(* IEC 61131-3 sources: daoli-st-library/DL_MathData (part 22) *)

(* ---- FC_DL_RealToUintSat.st ---- *)
(*
    FC_DL_RealToUintSat —— REAL 到 UINT 饱和防御转换
    ------------------------------------------------------------------
    分类      : DL_MathData / Convert
    前缀      : FC_DL_
    版本      : 1.0.0
    溯源      : IEC 61131-3 标准语义的道莅防御性实现
                （内部委托平台内建函数，外围统一错误码/钳位/双语文档；
                  未复制任何闭源厂商源码，参考实现仅限 MIT/Apache 许可）
    平台      : 纯 IEC 61131-3，CODESYS / TwinCAT / InoProShop 通用
    作者      : 道莅代码库 · PLC编程专家（R16）
    ------------------------------------------------------------------
    功能说明  : 将 REAL 输入防御性转换为 UINT 并作为返回值输出；
                非有限输入（NaN 或 ±INF）判为故障级 16#0001_0297，返回 0 且 bValid=FALSE；
                fIn < 0 时钳位至 0，置信息级 16#0001_01C6（UINT 无符号，负值不可表）；
                fIn 超出 UINT 上界 65535 时钳位至上界，置信息级 16#0001_01C7；
                钳位方向：下界 0 / 上界 65535（双侧饱和）；
                ±INF 采用平台安全幅值比较判定（阈值高于 REAL 最大有限值 3.402823E38），NaN 用 fIn <> fIn 自不等判定；
                域内转换委托平台内建 REAL_TO_UINT 语义，不重实现数学内核；
                信息级码属正常防御：bError=FALSE、bValid=TRUE，输出钳位后防御值。
    错误码    : 16#0001_0297 非有限输入（NaN 或 ±INF）——故障级，返回 0
                16#0001_01C6 负值输入，已钳位至 0——信息级，正常防御
                16#0001_01C7 输入超 UINT 上界，已钳位至 65535——信息级，正常防御
                16#0001_0298 预留禁用（故障级，不得挪用）
                16#0001_0299 预留禁用（故障级，不得挪用）
    状态机    : R6 标注 N/A —— 本组件为纯函数无顺序状态机，无 CASE 可写，非法状态不可能出现，故以本节说明替代 ELSE 兜底
    修订记录  : 2026-11-16 v1.0.0 首次入库（R16）
*)
FUNCTION FC_DL_RealToUintSat : UINT
VAR_INPUT
    fIn : REAL; // 待转换输入 [无量纲] / input value to convert
END_VAR
VAR_OUTPUT
    eErr   : UDINT; // 错误码，0=正常 / error id, 0=ok
    bError : BOOL;  // 是否出错，eErr 非 0 时为 TRUE / error flag, TRUE when eErr is nonzero
    bValid : BOOL;  // 输出是否有效可用 / output valid flag
END_VAR
VAR CONSTANT
    DL_UINT16_MAX     : LREAL := 65535.0; // UINT 域上界 65535，LREAL 承载 [无量纲] / UINT upper bound 65535 carried in LREAL
    DL_REAL_INF_GUARD : LREAL := 4.0E38;  // REAL 域 ±INF 判定阈值，高于 REAL 最大有限值 3.402823E38 [无量纲] / REAL +/-INF guard above max finite REAL 3.402823E38
END_VAR
VAR
    bNonFinite : BOOL; // 非有限（NaN 或 ±INF）判定结果 / non-finite (NaN or +/-INF) detection result
END_VAR

// 段 1｜返回值与错误状态预置 / segment 1, preset return value and error status
FC_DL_RealToUintSat := 0; // 故障缺省返回 0 [无量纲] / fault default returns 0
eErr   := 0;     // 预置无错误 / preset no error
bError := FALSE; // 预置无故障 / preset no fault
bValid := FALSE; // 预置无效，通过防御闸后置位 / preset invalid, set TRUE after guard passes

// 段 2｜非有限防御闸 / segment 2, non-finite guard
bNonFinite := (fIn <> fIn) OR (fIn > DL_REAL_INF_GUARD) OR (fIn < -DL_REAL_INF_GUARD); // NaN 自不等判定，±INF 用安全幅值比较 [无量纲] / NaN by self-inequality, +/-INF by safe magnitude compare
IF bNonFinite THEN
    FC_DL_RealToUintSat := 0; // 故障级返回 0 [无量纲] / fault level returns 0
    eErr   := 16#0001_0297;   // 非有限输入故障码 / non-finite input fault id
    bError := TRUE;           // 置故障标志 / set fault flag
    bValid := FALSE;          // 输出无效 / output invalid
    RETURN;                   // 立即返回 / immediate return
END_IF

// 段 3｜双侧饱和钳位与主体转换（末段） / segment 3, double-side saturating clamp and main conversion (final)
IF fIn < 0.0 THEN
    FC_DL_RealToUintSat := 0;  // 负值钳位至 0（UINT 无符号语义） / negative input clamped to 0 (UINT is unsigned)
    eErr := 16#0001_01C6;      // 信息级：负值已钳零 / info level: negative input clamped to zero
ELSIF fIn > DL_UINT16_MAX THEN
    FC_DL_RealToUintSat := 16#FFFF; // 正向钳位至 UINT 上界 65535 / clamp to UINT upper bound 65535
    eErr := 16#0001_01C7;           // 信息级：超上界已钳位 / info level: above upper bound, clamped
ELSE
    FC_DL_RealToUintSat := REAL_TO_UINT(fIn); // 域内委托平台内建 _TO_ 转换语义 / in-domain delegate to built-in _TO_ conversion
    eErr := 0; // 域内无错误 / in-domain, no error
END_IF
bError := FALSE; // 信息级钳位不置故障，故障分支已提前返回 / info-level clamp never raises fault, fault branch has returned
bValid := TRUE;  // 域内或钳位输出均有效可用 / in-domain or clamped output is valid
END_FUNCTION

(* ---- FC_DL_ReverseBitsWord.st ---- *)
(*==============================================================================
 * 组件名称 (Component)  : FC_DL_ReverseBitsWord
 * 所属子库 (Sublibrary) : DL_MathData
 * 归属目录 (Directory)  : C:\Library\DL_MathData
 * 当前版本 (Version)    : 1.0.0
 * 分类/来源标签         : 函数（FUNCTION）· 纯函数 · WORD 位反转与字节交换
 *                         iec-std-wrapper / bitstring
 * 兼容性   (Platform)   : CODESYS 3.5 / TwinCAT 3 / 汇川 InoProShop / 施耐德
 *                         Machine Expert；仅用 IEC 标准位运算 AND/OR/SHL/SHR
 * 溯源声明 (Provenance) : IEC 61131-3 标准语义的道莅防御性实现——内部委托平台标准库语义，
 *                         外围统一错误码 / 钳位 / 双语注释，严禁重实现数学内核。
 * 功能一句话 (Summary)  : WORD 全 16 位镜像反转（分治交换法）或字节序交换双模式，
 *                         服务 LSB-first CRC、LED 点阵与大小端报文适配。
 *
 * 功能描述 (Function)   : 位反转模式用四步分治交换（1 位组、2 位组、4 位组、
 *                         8 位组两两对换）实现全位镜像，无循环、无查表、常数时间；
 *                         字节交换模式一次完成高低字节对换；模式域外走 ELSE 兜底
 *                         回退位反转并报故障码，回文输入以信息级告知恒等结果。
 * 与既有件边界 (Boundary): 与 ShlEx/ShrEx 族正交——那些件做移位，本件做镜像；
 *                         平台内建 SWAP 指令非 IEC 标准，故字节交换同样手写实现。
 * 码位说明 (Codes)      : 信息 16#0002_3044 反转完成且结果回文（wOut 等于 wIn）
 *                         故障 16#0002_3045 模式域外，已回退位反转并照常输出
 *                         段 16#02_3_44~47，本件实占 44~45 两码。
 * 依赖说明 (Depends)    : 无 DL_ 内部依赖；零库函数依赖，纯 IEC 位运算符。
 * 红线自检 (Redline)    : 零全局依赖 ｜ 零 VAR_EXTERNAL ｜ 零 %I/%Q ｜ 纯 IEC 位运算
 *                         移位量 1/2/4/8 恒小于 16 位宽（归一达标）｜ 无除法面
 *                         ENUM 配 CASE 且 ELSE 兜底 ｜ 全变量双语同行注释
 * 修订历史 (Revision)   : 2026-11-18  v1.0.0  首版入库（R32 · 批 1）
 *============================================================================*)

FUNCTION FC_DL_ReverseBitsWord : BOOL
VAR_INPUT
    wIn   : WORD;                       // 源字 [位串] / Source word
    eMode : (eRevBits := 0, eRevBytes := 1);    // 模式枚举：全位反转或字节交换 / Mode enum: full bit reverse or byte swap
END_VAR
VAR_OUTPUT
    wOut    : WORD;                     // 反转结果 [位串] / Reversed result
    bPalin  : BOOL;                     // 回文标志，wOut 等于 wIn 时为真 / TRUE when the result equals the input
    uErrorId: UDINT;                    // 事件码，0 表示无事件 / Event code, zero means none
END_VAR
VAR
    w1 : WORD;    // 第一步交换结果（1 位组）[位串] / Stage one result, one-bit groups
    w2 : WORD;    // 第二步交换结果（2 位组）[位串] / Stage two result, two-bit groups
    w3 : WORD;    // 第三步交换结果（4 位组）[位串] / Stage three result, four-bit groups
    w4 : WORD;    // 第四步交换结果（8 位组，即全镜像）[位串] / Stage four result, full mirror
    uCode : UDINT; // 码位暂存，出口单点写入 [码] / Code staging
END_VAR

(* 段 1｜输出预置 / Pre-set *)
FC_DL_ReverseBitsWord := FALSE;
wOut    := 16#0000;
bPalin  := FALSE;
uErrorId := 16#0000_0000;
uCode   := 16#0000_0000;

(* 段 2｜模式分派（ENUM 配 CASE，ELSE 兜底拦截域外值）/ Mode dispatch with ELSE interception *)
CASE eMode OF

    eRevBits:
        (* 四步分治交换：相邻 1 位、2 位、4 位对换，最后高低 8 位整体对换
         * Four divide-and-conquer stages, constant time, no loop and no table *)
        w1 := ((wIn  AND 16#5555) SHL 1)  OR ((wIn  AND 16#AAAA) SHR 1);  // 相邻 1 位对换 / Adjacent one-bit swap
        w2 := ((w1   AND 16#3333) SHL 2)  OR ((w1   AND 16#CCCC) SHR 2);  // 相邻 2 位对换 / Adjacent two-bit swap
        w3 := ((w2   AND 16#0F0F) SHL 4)  OR ((w2   AND 16#F0F0) SHR 4);  // 相邻 4 位对换 / Adjacent four-bit swap
        w4 := ((w3   AND 16#00FF) SHL 8)  OR ((w3   AND 16#FF00) SHR 8);  // 高低 8 位对换，完成全镜像 / Final mirror
        wOut := w4;

    eRevBytes:
        (* 字节交换：低 8 位左移到高位，高 8 位右移到低位 / Swap the two bytes *)
        wOut := ((wIn AND 16#00FF) SHL 8) OR ((wIn AND 16#FF00) SHR 8);

ELSE
    (* 域外兜底：枚举被非法赋值（如强转越界）时回退位反转，绝不输出未定义值
     * Out-of-domain fallback: revert to bit reverse, never output an undefined value *)
    w1 := ((wIn  AND 16#5555) SHL 1)  OR ((wIn  AND 16#AAAA) SHR 1);
    w2 := ((w1   AND 16#3333) SHL 2)  OR ((w1   AND 16#CCCC) SHR 2);
    w3 := ((w2   AND 16#0F0F) SHL 4)  OR ((w2   AND 16#F0F0) SHR 4);
    w4 := ((w3   AND 16#00FF) SHL 8)  OR ((w3   AND 16#FF00) SHR 8);
    wOut := w4;
    uCode := 16#0002_3045;           // 故障级：模式域外已回退 / Fault: mode out of domain, reverted

END_CASE

(* 段 3｜回文告知与出口 / Palindrome notice and exit *)
IF wOut = wIn THEN
    bPalin := TRUE;                  // 恒等结果（回文字）告知 / Inform the identity result
    IF uCode = 16#0000_0000 THEN
        uCode := 16#0002_3044;       // 信息级：结果回文 / Info: palindromic result
    END_IF
END_IF
uErrorId := uCode;                   // 码位单点写入 / Single write point for the code
FC_DL_ReverseBitsWord := TRUE;
END_FUNCTION

(* ---- FC_DL_RmsCalc.st ---- *)
(*
    FC_DL_RmsCalc —— 窗口均方根（增量式平方累加防溢出 + 窗长钳位 + 非有限剔除）
    ------------------------------------------------------------------
    分类      : DL_MathData / Math-Statistics
    前缀      : FC_DL_
    版本      : 1.0.1
    来源标签  : iec-std-wrapper（T0）
    溯源      : IEC 61131-3 标准语义的道莅防御性实现
                （无状态纯函数，SQRT 为 IEC 标准内建；未复制任何闭源厂商源码）
    平台      : 纯 IEC 61131-3，CODESYS / TwinCAT / InoProShop 通用
    分工声明  : 与存量 FB_DL_SignalStatistics / FC_DL_StdDevOnline 分工——
                SignalStatistics 为驻留统计族（均值/方差多出口），StdDevOnline
                为在线流式标准差；本件为无状态数组窗口 RMS 单出口口径，
                与批 2 Safe 族惯性一致（无依赖，仅排期顺延）。
    作者      : 道莅代码库 · PLC 编程专家（R57）
    ------------------------------------------------------------------
    功能说明  : 对输入数组前 nCount 个样本求均方根。增量式累加 sum += x²/n
                防大数平方溢出（先除后加，边界十二）；窗长钳位 1..4096；
                非有限样本剔除并计数出口；有效样本数为零判错误返回 0。
    错误码    : 0000 正常 / 16#0003_0003 窗长已钳位 / 16#0003_0004 有效样本为零
                / 16#0003_0005 非有限样本已剔除（信息级，bValid 保持 TRUE）
    bValid 偏离段: 部分剔除时 bValid 保持 TRUE——有效样本统计量仍可用（与
                0303 钳位件 bValid=FALSE 的口径差异在此声明，v1.0.1）。
    修订记录  : 2026-11-21 v1.0.0 首次入库（R57 批 3 · 序号 12）
                2026-11-21 v1.0.1 R58 返修：部分剔除（nUsed>0 且 nNanCnt>0）
                置信息级 0003_0005（首事件闸），调用方可感知口径已收窄；
                全剔除路径 0304 优先级在先不动。
*)
FUNCTION FC_DL_RmsCalc : LREAL
VAR_IN_OUT
    afData : ARRAY[0..4095] OF LREAL; // 样本数组 [工程单位]，前 nCount 个有效 / the sample array, the first nCount entries valid
END_VAR
VAR_INPUT
    nCount : DINT; // 样本数 [个]，钳位 1..4096 / the sample count, clamped to one through four thousand ninety six
END_VAR
VAR_OUTPUT
    eErr     : UDINT; // 错误码，0 = 正常 / error code, zero is ok
    bError   : BOOL;  // 出错标志，eErr 非 0 时为真 / error flag, true when eErr is nonzero
    bValid   : BOOL;  // 结果是否为真实值，钳位/剔除降级时可能为假 / the result is the true value, false when degraded
    nNanCnt  : UDINT; // 剔除的非有限样本数 [个] / the excluded non finite sample count
END_VAR
VAR
    nI     : DINT;  // 循环计数 [个] / the loop counter
    nUsed  : DINT;  // 实际参与样本数 [个] / the actually used sample count
    lrSum  : LREAL; // 增量式平方和 [工程单位平方] / the incremental sum of squares
    lrX    : LREAL; // 当前样本 [工程单位] / the current sample [engineering unit]
    bClamp : BOOL;  // 窗长钳位发生 [-] / a window clamp happened
END_VAR
VAR CONSTANT
    DL_RMS_NMAX : DINT := 4096; // 窗长上限 [个]，与数组容量一致 / the window bound, aligned with the array capacity
END_VAR

// 段 1｜返回值与错误状态预置安全值（四段式第一段，R45）/ segment 1, preset the return and error states
FC_DL_RmsCalc := 0.0; // 返回值预置安全值 0.0 / preset the return to the safe zero
eErr   := 16#0000_0000; // 错误码预置正常 / preset the code to ok
bError := FALSE; // 错误标志预置假 / preset the error flag false
bValid := TRUE; // 有效标志预置真 / preset the valid flag true
nNanCnt := 0; // 剔除计数预置零 / preset the excluded count zero
bClamp := FALSE; // 钳位标志预置假 / preset the clamp flag false

// 段 2｜窗长钳位 1..4096（边界十二；上界与数组容量一致，索引结构性安全）/ segment 2, the window clamp
IF nCount < 1 THEN // 低于下界 / below the floor
    nCount := 1; // 钳到 1 / clamp to one
    bClamp := TRUE; // 置钳位标记 / raise the clamp flag
ELSIF nCount > DL_RMS_NMAX THEN // 高于上界 / above the bound
    nCount := DL_RMS_NMAX; // 钳到上限 / clamp to the bound
    bClamp := TRUE; // 置钳位标记 / raise the clamp flag
END_IF
IF bClamp THEN // 钳位发生时置信息级 / raise the informational code on a clamp
    eErr   := 16#0003_0003; // 信息级：窗长已钳位 / informational, the window clamped
    bError := TRUE; // 置错误标志 / raise the error flag
    bValid := FALSE; // 钳位口径非原始窗长口径 / the clamped window is not the requested one
END_IF

// 段 3｜增量式平方累加：sum += x²/n（先除后加防大数溢出，边界十二）/ segment 3, the incremental accumulation
lrSum := 0.0; // 平方和清零 / clear the sum
nUsed := 0; // 参与样本数清零 / clear the used count
FOR nI := 0 TO nCount - 1 DO // 有界循环（nCount 已钳 ≤4096）/ the bounded loop
    lrX := afData[nI]; // 取样本（索引已证在数组界内）/ take the sample, the index proven inside the bounds
    IF (lrX = lrX) AND ((lrX - lrX) = (lrX - lrX)) THEN // 非有限双判据通过才参与 / only finite samples participate
        lrSum := lrSum + lrX * lrX / INT_TO_LREAL(nCount); // 先除窗长再加，防 x² 大数溢出 / divide first then add against overflow
        nUsed := nUsed + 1; // 参与计数推进 / advance the used count
    ELSE // 非有限样本剔除 / a non finite sample excluded
        nNanCnt := nNanCnt + 1; // 剔除计数推进 / advance the excluded count
    END_IF
END_FOR

// 段 3b｜部分剔除信息级置码（v1.0.1：首事件闸，0303 先发则不再覆盖）/ segment 3b, the partial exclusion informational code
IF (nNanCnt > 0) AND (nUsed > 0) AND (eErr = 16#0000_0000) THEN // 部分剔除且无先发事件 / a partial exclusion with no earlier event
    eErr   := 16#0003_0005; // 信息级：非有限样本已剔除，口径为有效样本 RMS / informational, non finite samples excluded, the effective sample RMS
    bError := TRUE; // 置错误标志（信息级随事件置位惯例）/ raise the error flag
END_IF // bValid 保持 TRUE：有效样本统计量仍可用（头注释偏离段声明）/ bValid stays true, the effective sample statistic remains usable

// 段 4｜结果计算与兜底 / segment 4, the result and the guard
IF nUsed > 0 THEN // 有有效样本 / with valid samples
    FC_DL_RmsCalc := SQRT(lrSum * INT_TO_LREAL(nCount) / INT_TO_LREAL(nUsed)); // 复原除子后开方（除子已证大于零）/ restore the divisor then the square root
ELSE // 全部剔除 / all excluded
    eErr   := 16#0003_0004; // 错误级：有效样本为零 / error grade, no valid sample
    bError := TRUE; // 置错误标志 / raise the error flag
    bValid := FALSE; // 输出不可用 / the output void
END_IF
IF (FC_DL_RmsCalc <> FC_DL_RmsCalc) OR ((FC_DL_RmsCalc - FC_DL_RmsCalc) <> (FC_DL_RmsCalc - FC_DL_RmsCalc)) THEN // 结果非有限兜底 / the non finite result guard
    FC_DL_RmsCalc := 0.0; // 兜底安全值 / the bottom-line safe value
    bValid := FALSE; // 输出不可用 / the output void
END_IF
END_FUNCTION

(* ---- FC_DL_RoundBankEx.st ---- *)
(*
    FC_DL_RoundBankEx —— ROUND 明确口径包装（银行家/半进可选，LREAL 域）
    ------------------------------------------------------------------
    分类      : DL_MathData / Rounding
    前缀      : FC_DL_
    版本      : 1.0.0
    溯源      : IEC 61131-3 标准语义的道莅防御性实现
                （内部委托 TRUNC 标准函数与比较语义，外围统一错误码/钳位/双语文档；
                  未复制任何闭源厂商源码，参考实现仅限 MIT/Apache 许可）
    平台      : 纯 IEC 61131-3，CODESYS / TwinCAT / InoProShop 通用
    作者      : 道莅代码库 · PLC编程专家（R40）
    ------------------------------------------------------------------
    功能说明  : 将 fIn 舍入到最近整数（仍以 LREAL 返回），0.5 进位方向全平台
                显式统一，杜绝 ROUND 内建在三平台的半进/半退差异泄漏：
                bHalfUp = FALSE（缺省）：0.5 进位到最近的偶数（银行家口径）；
                bHalfUp = TRUE：0.5 一律进位（向远离零方向，半进口径）；
                非半点小数一律按最近整数舍入（>0.5 进、<0.5 退）；
                非有限输入（NaN 或 ±Inf）判为故障级 16#0001_03CF，返回 0.0 且
                bValid=FALSE（NaN 参与舍入在三平台行为不一致，一律拦截）；
                超整数分辨率恒等直通：|fIn| ≥ 2^53（9.007199254740992E15）时
                该幅值下 LREAL 相邻可表数间距已大于 1，输入必为整数值，
                舍入恒等直通并置信息级 16#0001_0496；
                溢出面分析（R63 反算句）：|fIn| < 2^53 时结果 |fRnd| ≤ |fIn| + 1 ≤ 2^53，
                恒在 LREAL 可表域内，无溢出路径，无需饱和钳位（算法已证）；
                半点检测口径：ABS(fFrac − 0.5) < 1.0E-9 视为半点（差值在 1E-9 内的
                近半点值按半点口径处理，取舍显式化，避免浮点表示误差致半点漏判）。
    错误码    : 16#0001_03CF 任一输入非有限（NaN 或 ±Inf）——故障级，返回 0.0
                16#0001_0496 输入幅值 ≥ 2^53，超整数分辨率，恒等直通——信息级，正常防御
                （R90 反证句：恒等直通场景无法由返回值观测——直通值与舍入结果同为
                  合法整数值，bValid=TRUE 组合相同，现有输出无法还原「分辨率已耗尽」
                  事实，故占信息码）
    状态机    : R6 标注 N/A —— 本组件为纯函数无顺序状态机，无 CASE 可写，
                非法状态不可能出现，故以本节说明替代 ELSE 兜底
    修订记录  : 2026-11-19 v1.0.0 首次入库（R40 · 批 2 · T0 快车道）
*)
FUNCTION FC_DL_RoundBankEx : LREAL
VAR_INPUT
    fIn     : LREAL;         // 待舍入输入 [无量纲] ｜ input to round
    bHalfUp : BOOL := FALSE; // 半点口径，FALSE=进位到最近偶数（银行家），TRUE=一律半进 ｜ half-point mode, FALSE=round half to even (banker's), TRUE=round half away from zero
END_VAR
VAR_OUTPUT
    eErr   : UDINT; // 错误码，0=正常，16#0001_04XX=信息级，16#0001_03XX=故障级 ｜ error id, 0=ok, 16#0001_04XX=info, 16#0001_03XX=fault
    bError : BOOL;  // 是否出错，eErr 落故障级时为 TRUE ｜ fault flag, TRUE when eErr is fault level
    bValid : BOOL;  // 输出是否有效可用 ｜ output valid flag
END_VAR
VAR CONSTANT
    DL_ROUND_ID_LIMIT : LREAL := 9.007199254740992E15; // 恒等直通幅值限 = 2^53 [无量纲] ｜ identity pass-through magnitude limit = 2^53
    DL_ROUND_HALF     : LREAL := 0.5;                  // 半点判据常数 [无量纲] ｜ half-point constant
    DL_ROUND_TOL      : LREAL := 1.0E-9;               // 半点检测容差 [无量纲] ｜ half-point detection tolerance
    DL_ROUND_ONE      : LREAL := 1.0;                  // 进位步长 [无量纲] ｜ carry step
    DL_ROUND_TWO      : LREAL := 2.0;                  // 偶数判定基数 [无量纲] ｜ even-test radix
END_VAR
VAR
    bNonFinite : BOOL;  // 非有限（NaN 或 ±Inf）判定结果 ｜ non-finite (NaN or +/-Inf) detection result
    fAbs       : LREAL; // 输入绝对值 [无量纲] ｜ absolute value of the input
    fInt       : LREAL; // 绝对值的整数部分（TRUNC 向零截断）[无量纲] ｜ integer part of the magnitude (TRUNC toward zero)
    fFrac      : LREAL; // 绝对值的小数部分 [无量纲] ｜ fractional part of the magnitude
    fRnd       : LREAL; // 舍入后的绝对值结果 [无量纲] ｜ rounded magnitude result
END_VAR

// 段 1｜返回值与错误状态预置 ｜ segment 1, preset return value and error status
FC_DL_RoundBankEx := 0.0; // 故障缺省返回 0 [无量纲] ｜ fault default returns 0
eErr   := 0;     // 预置无错误 ｜ preset no error
bError := FALSE; // 预置无故障 ｜ preset no fault
bValid := FALSE; // 预置无效，通过防御闸后置位 ｜ preset invalid, set TRUE after guard passes

// 段 2｜非有限防御闸（早退） ｜ segment 2, non-finite guard (early return)
bNonFinite := (fIn <> fIn) OR ((fIn - fIn) <> (fIn - fIn)); // NaN 自不等 + 差值自减判 ±Inf [无量纲] ｜ NaN by self-inequality, +/-Inf by self-subtraction
IF bNonFinite THEN
    FC_DL_RoundBankEx := 0.0; // 故障级返回 0 [无量纲] ｜ fault level returns 0
    eErr   := 16#0001_03CF;   // 非有限输入故障码 ｜ non-finite input fault id
    bError := TRUE;           // 置故障标志（R45 配对）｜ raise the fault flag (R45 pairing)
    bValid := FALSE;          // 输出无效 ｜ output invalid
    RETURN;                   // 早退 ｜ early return
END_IF

// 段 3｜超整数分辨率恒等直通（信息级） ｜ segment 3, identity pass-through beyond integer resolution (info level)
IF ABS(fIn) >= DL_ROUND_ID_LIMIT THEN
    FC_DL_RoundBankEx := fIn; // 分辨率耗尽，舍入恒等直通 [无量纲] ｜ resolution exhausted, rounding is identity
    eErr   := 16#0001_0496;   // 信息级：超分辨率恒等直通 ｜ info level: identity pass-through beyond resolution
    bError := FALSE;          // 信息级不置故障 ｜ info level raises no fault
    bValid := TRUE;           // 直通输出有效 ｜ pass-through output is valid
    RETURN;                   // 早退 ｜ early return
END_IF

// 段 4｜绝对域分解与舍入主体（末段） ｜ segment 4, magnitude decomposition and rounding body (final)
fAbs  := ABS(fIn);        // 取绝对值 [无量纲] ｜ take the magnitude
fInt  := TRUNC(fAbs);     // 整数部分（TRUNC 向零截断，绝对域恒非负）｜ integer part (TRUNC toward zero, non-negative in magnitude domain)
fFrac := fAbs - fInt;     // 小数部分（fInt ≥ fAbs/2 或 fInt=0，减法在 2^53 内精确，无消去误差）｜ fractional part (subtraction exact below 2^53, no cancellation error)
IF ABS(fFrac - DL_ROUND_HALF) < DL_ROUND_TOL THEN
    // 半点口径：按 bHalfUp 显式分流 ｜ half-point mode: explicit branch by bHalfUp
    IF bHalfUp THEN
        fRnd := fInt + DL_ROUND_ONE;  // 半进口径：一律进位（远离零）｜ half-up mode: always carry (away from zero)
    ELSE
        // 银行家口径：进位到最近偶数（偶数判定用差值容差比较，禁浮点直等）｜ banker's mode: round half to even (even test by difference tolerance, no direct float equality)
        IF ABS(fInt - DL_ROUND_TWO * TRUNC(fInt / DL_ROUND_TWO)) < DL_ROUND_TOL THEN
            fRnd := fInt;                 // 整数部分为偶，退位保持 ｜ integer part even, keep it
        ELSE
            fRnd := fInt + DL_ROUND_ONE;  // 整数部分为奇，进位到偶 ｜ integer part odd, carry to even
        END_IF
    END_IF
ELSIF fFrac > DL_ROUND_HALF THEN
    fRnd := fInt + DL_ROUND_ONE;  // 非半点且大于半点，进位 ｜ beyond the half-point, carry
ELSE
    fRnd := fInt;                 // 非半点且小于半点，退位 ｜ below the half-point, keep
END_IF

// 段 5｜出口装配：恢复符号并单点写出 ｜ segment 5, exit assembly: restore the sign and write once
IF fIn < 0.0 THEN
    FC_DL_RoundBankEx := -fRnd; // 负输入恢复负号 [无量纲] ｜ negative input restores the sign
ELSE
    FC_DL_RoundBankEx := fRnd;  // 非负输入直通 [无量纲] ｜ non-negative input passes through
END_IF
bError := FALSE; // 正常出口不置故障 ｜ normal exit raises no fault
bValid := TRUE;  // 舍入输出有效可用 ｜ rounding output is valid
END_FUNCTION

(* ---- FC_DL_RoundSat.st ---- *)
(*==============================================================================
 * 组件名称 (Component)  : FC_DL_RoundSat
 * 所属子库 (Sublibrary) : DL_MathData
 * 当前版本 (Version)    : 1.0.0
 * 兼容性   (Platform)   : CODESYS 3.5 / TwinCAT 3 / 汇川 InoProShop / Machine Expert
 *                         仅依赖 Standard.library 的 ROUND / ABS 内建函数，
 *                         不重实现取整内核，无厂商数学方言依赖
 * 功能一句话 (Summary)  : 四舍五入取整饱和包装：非有限拦截 + DINT 越界
 *                         钳到端点不回绕，半值取向写死为「四舍五入远离零」。
 * 功能描述 (Function)   : 对输入实数 fX 四舍五入取整为 DINT。闸门次序写死：
 *                         ① 非有限复检先行（NaN 用 x <> x 判据、无穷用
 *                         ABS(x) 超有限性上界判据），命中返回 0 + 故障码；
 *                         ② DINT 越界饱和闸——fX >= 2147483647.5 时 ROUND
 *                         必溢出，钳到 DINT 上端点 2147483647 并置信息码；
 *                         fX <= -2147483648.5 时钳到下端点 -2147483648
 *                         并置信息码，绝不回绕；③ 域内委托内建 ROUND。
 * 溯源     (Origin)     : IEC 61131-3 标准语义的道莅防御性实现
 *                         （接口语义由 IEC 61131-3 定义，clean-room 重写，
 *                         参考公开标准条款）
 * 半值取向 (Half Policy): 「.5 半值取向」写死为本库取「四舍五入远离零」
 *                         （round half away from zero，多数平台 ROUND 语义）；
 *                         需要银行家舍入（round half to even）的调用方用
 *                         FLOOR / CEIL / TRUNC 组合自行复现，本件不提供。
 * 码位     (Diag Codes) : 故障级 16#0001_022B（本件独占）：
 *                           输入非有限（NaN / 无穷），返回 0；
 *                         信息级 16#0001_015B（本件独占）：
 *                           DINT 越界已钳位到端点（上端点或下端点，
 *                           饱和是正常防御行为，不回绕）。
 * 类型裁定 (Type Note)  : 码位段 16#0001_xxxx 为全库共享 32 位段，WORD 容量不足，
 *                         故 eErr 采用 UDINT 承载（与库内 uErrorId : UDINT 惯例
 *                         一致，沿 R14 批 3 同一裁定）。
 * 依赖     (Depends)    : 无 DL_ 内部依赖；Standard.library: ROUND / ABS
 * 红线自检 (Redline)    : R1 ✓ 零全局变量与外部变量引用 ｜ R2 ✓ 零物理 IO 地址直写
 *                         R3 ✓ 纯 IEC 61131-3 ｜ R4 ✓ 非有限拦截 + 越界饱和不回绕
 *                         R5 ✓ 全变量中英双语同行注释
 *                         R6 N/A（纯函数，无 CASE/ENUM 状态机，按批 4 口径标 N/A）
 *                         R7 N/A（FC 为纯函数，无实例调用，头注释显式说明）
 * 防御行为声明 (Defense): ① 非有限复检先行：NaN 判据 fX <> fX（NaN 与任何值
 *                           包括自身比较均为不等，库内既有写法）、无穷判据
 *                           ABS(fX) > 1.0E308，命中即不调内建、早退返回 0；
 *                         ② 饱和阈值取 2147483647.5 / -2147483648.5（而非
 *                           DINT 端点本身）：|x| <= 2^53 内 LREAL 可精确表示
 *                           该阈值，ROUND 在阈值内侧（不含）结果必落在
 *                           [DINT_MIN, DINT_MAX]，阈值及外侧一律钳端点置码，
 *                           绝不回绕（与平台整数回绕行为的差异点）；
 *                         ③ 域内委托内建 ROUND 内核（四舍五入远离零），
 *                           本件不重实现取整；
 *                         ④ 饱和是显式信息码 16#0001_015B，不是静默钳位，
 *                           现场可凭码定位「量纲/增益配错导致的巨数」；
 *                         ⑤ 阈值与端点、1.0E308 有限性上界均提为只读常量，
 *                           禁魔法数；
 *                         ⑥ 浮点全程不用等号直比判数值相等，仅用 < > 与
 *                           NaN 自不等判据，符合浮点容差红线口径。
 * 修订历史 (Revision)   :
 *   2026-11-16  v1.0.0  首版入库（R14 批 4 · T0 快车道）
 *============================================================================*)
FUNCTION FC_DL_RoundSat : DINT
VAR_INPUT
    fX : LREAL; // 输入实数 [无量纲] / Input real value [dimensionless]
END_VAR
VAR_OUTPUT
    eErr : UDINT; // 错误码，16#0001_022B=非有限输入，16#0001_015B=越界钳位到 DINT 端点，0=无事件 / Error code, 16#0001_022B=non-finite input, 16#0001_015B=clamped to a DINT endpoint, 0=no event
END_VAR
VAR CONSTANT
    DL_RND_FINITE : LREAL := 1.0E308;       // 有限性上界 [无量纲]，超界判无穷（库内既有写法）/ Finiteness bound, values beyond treated as infinity (library idiom)
    DL_RND_HI     : LREAL := 2147483647.5;  // 饱和上阈 [无量纲]，fX >= 此值 ROUND 必溢出上端点 / Saturation upper threshold, ROUND overflows above it
    DL_RND_LO     : LREAL := -2147483648.5; // 饱和下阈 [无量纲]，fX <= 此值 ROUND 必溢出下端点 / Saturation lower threshold, ROUND overflows below it
    DL_RND_DMAX   : DINT  := 2147483647;    // DINT 上端点 [个]，钳位目标 / DINT upper endpoint, clamping target
    DL_RND_DMIN   : DINT  := -2147483648;   // DINT 下端点 [个]，钳位目标 / DINT lower endpoint, clamping target
END_VAR

(*------------------------------------------------------------------------------
 * 段 1｜返回值与错误码预置：先归零，任何早退路径都不会留下脏码
 *      Preset return value and error code so no early-exit path leaves a stale code
 *-----------------------------------------------------------------------------*)
FC_DL_RoundSat := 0;           // 返回值预置 0 [个] / Preset return value to zero
eErr           := 16#0000_0000;   // 错误码预置无事件 / Preset error code to no event

(*------------------------------------------------------------------------------
 * 段 2｜非有限复检先行（防御声明①）：NaN / 无穷一律不进内建内核
 *      Non-finite recheck first (defense note 1): NaN and infinity never reach
 *      the built-in kernel
 *-----------------------------------------------------------------------------*)
IF (fX <> fX) OR (ABS(fX) > DL_RND_FINITE) THEN
    eErr := 16#0001_022B;   // 故障码：输入非有限（NaN / 无穷），返回 0 / Fault: non-finite input (NaN or infinity), zero returned
    RETURN;                 // 返回预置值 0 [个] / Return preset value zero
END_IF

(*------------------------------------------------------------------------------
 * 段 3｜DINT 越界饱和闸（防御声明②④）：越界钳到端点并置信息码，
 *      绝不回绕；上/下端点对称处理
 *      DINT out-of-range saturation gate (defense notes 2 and 4): clamp to the
 *      endpoint with an informational code, never wrap; symmetric up and down
 *-----------------------------------------------------------------------------*)
IF fX >= DL_RND_HI THEN
    FC_DL_RoundSat := DL_RND_DMAX;   // 钳到 DINT 上端点 2147483647 [个] / Clamp to the DINT upper endpoint
    eErr := 16#0001_015B;            // 信息码：越界已钳位到上端点（不回绕）/ Informational: clamped to the upper endpoint, no wrap
    RETURN;                          // 饱和早退，不进内建 / Saturating early exit, built-in not called
END_IF

IF fX <= DL_RND_LO THEN
    FC_DL_RoundSat := DL_RND_DMIN;   // 钳到 DINT 下端点 -2147483648 [个] / Clamp to the DINT lower endpoint
    eErr := 16#0001_015B;            // 信息码：越界已钳位到下端点（不回绕）/ Informational: clamped to the lower endpoint, no wrap
    RETURN;                          // 饱和早退，不进内建 / Saturating early exit, built-in not called
END_IF

(*------------------------------------------------------------------------------
 * 段 4｜域内委托内建内核（防御声明③）：阈值内侧必落在 DINT 域，
 *      委托内建 ROUND（四舍五入远离零，半值取向见头注释）
 *      In-domain delegation to the built-in kernel (defense note 3): inside
 *      the thresholds the result always fits DINT, delegate to the built-in
 *      ROUND (round half away from zero, see the half policy in the header)
 *-----------------------------------------------------------------------------*)
FC_DL_RoundSat := ROUND(fX);   // 委托内建 ROUND 内核，不自实现取整 / Delegate to the built-in ROUND kernel, no re-implementation
END_FUNCTION

(* ---- FC_DL_RoundSigFigs.st ---- *)
(*
  ==================================================================
  组件名 Component  : FC_DL_RoundSigFigs
  分类   Category   : DL_MathData
  复杂度 Complexity  : cx3
  版本   Version    : 1.0.0
  功能   Purpose    : 按有效数字位数舍入。把 fVal 舍入到 nSigFigs 位有效数字
                      （半值远离零），10 的幂用整数循环累乘实现（禁 ** 幂运算符）；
                      nSigFigs 越域回钳 1..15 并置 bClamped，非有限值透传并置
                      bInvalid，舍入位置超出 DINT 安全域时原值透传并置 bClamped。
  来源   Source     : t2-1-lgf-math
  溯源   Origin     : IEC 61131-3 标准语义的道莅防御性实现；有效数字舍入为公开数值
                      方法，clean-room 自研实现，未复制任何闭源代码行。
  平台   Platform   : 纯 IEC 61131-3（LREAL / TRUNC / 循环累乘，无私有库、无幂运算符）
  作者   Author     : 道莅代码库 · PLC 编程专家（R56）
  ------------------------------------------------------------------
  边界 Boundary     :
                      一 本件只做十进制有效位舍入，不做定点小数位舍入（属主边界）；
                      二 DINT 可表上界反算（R63）：DINT 上限 2.147E9，取 1.0E9 为
                         TRUNC 安全阈；被舍整数部分 q >= 1.0E9 时（即 nSigFigs >= 10
                         且量级 >= 1E9），拆高低两段各 TRUNC（每段 < 1.0E9 可表），
                         合成值 < 1E15 < 2^53 在 LREAL 精确可表；
                      三 指数域钳 [-300, 300]：LREAL 上限 1.797E308，10^308 可表、
                         10^309 不可表；越钳透传原值并置 bClamped；
                      四 非有限输入透传（规格明示方向）并置 bInvalid，不参与舍入；
                      五 无全局变量、无外部变量声明、无物理地址寻址、无定时器（纯函数）。
  输出契约 Output contract:
                      fOut 在 bInvalid = FALSE 时为舍入结果，bInvalid = TRUE 时透传 fVal；
                      本件为纯函数，无跨扫描周期状态驻留。
  修订记录 Revision  :
    2026-11-20  v1.0.0  R56 首版（批 1 · 序号 3）
  ==================================================================
*)

FUNCTION FC_DL_RoundSigFigs : BOOL
VAR_INPUT
    fVal     : LREAL; // 待舍入值（带符号）[工程单位] / the value to be rounded, signed [engineering unit]
    nSigFigs : INT;   // 有效数字位数，越域回钳 1..15 [位] / significant digit count, clamped one through fifteen [digit]
END_VAR
VAR_OUTPUT
    fOut     : LREAL; // 舍入结果（带符号）[工程单位] / the rounded result, signed [engineering unit]
    bInvalid : BOOL;  // 非有限输入透传标志 [-] / the passthrough flag for a non finite input
    bClamped : BOOL;  // 位数或指数被回钳标志 [-] / the clamp flag for the digit count or the exponent
END_VAR
VAR
    _nSig    : INT := 1;    // 钳定后的有效位数 [位] / the clamped significant digit count [digit]
    _fAbs    : LREAL := 0.0;  // 绝对值工作值 [工程单位] / absolute value working quantity
    _fV      : LREAL := 0.0;  // 量级归一工作值 [工程单位] / magnitude normalising working quantity
    _eDec    : DINT := 0;     // 十进位阶（最高位有效数字所在幂）[幂] / decimal decade exponent of the leading digit
    _nPow    : DINT := 0;     // 舍入位置的十的幂（10^nPow）[幂] / power of ten at the rounding position
    _fP      : LREAL := 1.0;  // 十的幂累乘值 [无量纲] / accumulated power of ten
    _fQ      : LREAL := 0.0;  // 被舍实数（|fVal| / 10^nPow）[无量纲] / the value to be rounded integrally
    _fQHi    : LREAL := 0.0;  // 高段被舍实数 [无量纲] / the high segment to be rounded
    _fQLo    : LREAL := 0.0;  // 低段被舍实数 [无量纲] / the low segment to be rounded
    _nHi     : DINT := 0;     // 高段整数部分 [无量纲] / the high segment integer part
    _nLo     : DINT := 0;     // 低段整数部分 [无量纲] / the low segment integer part
    _fR      : LREAL := 0.0;  // 舍入后的整数（LREAL 精确表出）[无量纲] / the rounded integer, exactly representable in LREAL
    _i       : DINT := 0;     // 累乘循环游标 [次] / accumulation loop cursor
END_VAR

// 段 1｜非有限闸：透传并置标志（规格明示透传方向）/ segment 1, finiteness gate, passthrough per the specification
bInvalid := (fVal <> fVal) OR ((fVal - fVal) <> (fVal - fVal)); // NaN 自反、Inf 差值自减 / NaN by reflexivity, Inf by the self difference
IF bInvalid THEN // 非有限输入 / non finite input
    fOut := fVal; // 透传（规格明示）/ passthrough per the specification
    bClamped := FALSE; // 钳位标志不成立 / the clamp flag is false
    FC_DL_RoundSigFigs := FALSE; // 函数返回失败 / the function returns failure
    RETURN; // 早退 / early return
END_IF
bInvalid := FALSE; // 有限输入，标志不成立 / finite input, the flag is false
bClamped := FALSE; // 钳位标志预置假 / preset the clamp flag to false
FC_DL_RoundSigFigs := TRUE; // 默认返回成功 / default to success

// 段 2｜位数回钳 1..15（R117 两级回退：一级常量钳定）/ segment 2, digit count clamp
_nSig := nSigFigs; // 位数直通 / the count passes through
IF _nSig < 1 THEN // 下越域 / below the floor
    _nSig := 1; // 回钳到一位 / clamp to one digit
    bClamped := TRUE; // 置钳位标志 / raise the clamp flag
ELSIF _nSig > 15 THEN // 上越域 / above the ceiling
    _nSig := 15; // 回钳到十五位 / clamp to fifteen digits
    bClamped := TRUE; // 置钳位标志 / raise the clamp flag
END_IF

// 段 3｜零值与超小值快速出口 / segment 3, the fast exits for zero and tiny magnitudes
_fAbs := ABS(fVal); // 绝对值 / the absolute value
IF _fAbs < 1.0E-300 THEN // 量级低于指数域下限，舍入无意义 / the magnitude is below the exponent floor
    fOut := fVal; // 原值透传 / the value passes through
    RETURN; // 早退 / early return
END_IF

// 段 4｜十进位阶定位：整数循环归一（禁 **）/ segment 4, decade location by integer loops
_fV := _fAbs; // 归一工作值起步 / start the normalising working value
_eDec := 0; // 位阶清零 / clear the decade exponent
WHILE (_fV >= 10.0) AND (_eDec < 320) DO // 向上归一到 [1, 10) / normalise upward into the unit decade
    _fV := _fV / 10.0; // 除十 / divide by ten
    _eDec := _eDec + 1; // 位阶递增 / increment the decade
END_WHILE
WHILE (_fV < 1.0) AND (_eDec > -320) DO // 向下归一到 [1, 10) / normalise downward into the unit decade
    _fV := _fV * 10.0; // 乘十 / multiply by ten
    _eDec := _eDec - 1; // 位阶递减 / decrement the decade
END_WHILE

// 段 5｜舍入位置的十的幂：nPow = eDec - (nSig - 1)，越域钳 [-300, 300] / segment 5, the power at the rounding position
_nPow := _eDec - INT_TO_DINT(_nSig) + 1; // 目标幂（用钳定后位数）/ the target power from the clamped count
IF _nPow < -300 THEN // 下越域（10^-301 不可表）/ below the representable floor
    _nPow := -300; // 回钳 / clamp
    bClamped := TRUE; // 置钳位标志 / raise the clamp flag
ELSIF _nPow > 300 THEN // 上越域（10^301 不可表，R63 反算）/ above the representable ceiling
    _nPow := 300; // 回钳 / clamp
    bClamped := TRUE; // 置钳位标志 / raise the clamp flag
END_IF
_fP := 1.0; // 累乘起步一 / start the accumulation at one
IF _nPow >= 0 THEN // 正幂累乘 / the positive accumulation
    _i := 0; // 游标清零 / clear the cursor
    WHILE _i < _nPow DO // 累乘到目标幂 / accumulate to the target power
        _fP := _fP * 10.0; // 乘十 / multiply by ten
        _i := _i + 1; // 游标递增 / increment the cursor
    END_WHILE
ELSE // 负幂累乘 / the negative accumulation
    _i := 0; // 游标清零 / clear the cursor
    WHILE _i > _nPow DO // 累乘到目标幂 / accumulate to the target power
        _fP := _fP / 10.0; // 除十 / divide by ten
        _i := _i - 1; // 游标递减 / decrement the cursor
    END_WHILE
END_IF

// 段 6｜被舍实数与两段舍入（DINT 可表性分段，R63）/ segment 6, the value to be rounded and the two segment rounding
_fQ := _fAbs / _fP; // 被舍实数，除子为累乘幂已证非零 / the value to be rounded, the divisor is the proven power
IF _fQ < 1.0E9 THEN // 单段安全：q < 1.0E9 < DINT 上限（R63 反算）/ single segment safe against the DINT ceiling
    _nLo := TRUNC(_fQ + 0.5); // 半值远离零的整数舍入（|fVal| 口径恒正）/ integral rounding half away from zero on the always positive magnitude
    _fR := DINT_TO_LREAL(_nLo); // 整数精确落 LREAL / the integer lands exactly in LREAL
ELSE // 两段分解：高段 < 1.0E9、低段 < 1.0E6 均可表 / the two segment decomposition, both segments representable
    _fQHi := _fQ / 1000000.0; // 高段 = q / 1E6 / the high segment
    _nHi := TRUNC(_fQHi); // 高段截断 / truncate the high segment
    _fQLo := _fQ - DINT_TO_LREAL(_nHi) * 1000000.0; // 低段 = 余量 / the low segment remainder
    _nLo := TRUNC(_fQLo + 0.5); // 低段舍入 / round the low segment
    _fR := DINT_TO_LREAL(_nHi) * 1000000.0 + DINT_TO_LREAL(_nLo); // 合成（< 1E15 < 2^53 精确，进位由加法自然承载）/ the composition, exact below two to the fifty third, the carry rides the addition
END_IF

// 段 7｜符号回贴与出口 / segment 7, sign restore and the outlet
IF fVal < 0.0 THEN // 负值 / a negative value
    fOut := -_fR * _fP; // 符号回贴 / restore the sign
ELSE // 非负值 / a non negative value
    fOut := _fR * _fP; // 直接过出口 / straight to the outlet
END_IF
END_FUNCTION

(* ---- FC_DL_RoundToMultipleInt.st ---- *)
(*==============================================================================
 * 组件名称 : FC_DL_RoundToMultipleInt ｜ 子库 : DL_MathData ｜ v1.0.1 ｜ 2026-11-24
 * 平台     : CODESYS 3.5 / TwinCAT 3 / InoProShop / Machine Expert（纯 IEC，无厂商库）
 * 功能简介 : 整数四舍五入到 nMultiple 的最近倍数（半值远离零舍入，
 *            Round Half Away From Zero）。纯整数算术实现，先向零截断得
 *            基准倍数，再按"余量是否过半"进位 / 退位，无浮点精度损失。
 * 契约     : 返回四舍五入后的倍数值；nMultiple <= 0 恒返回 0 并置 bError；
 *            纯函数无状态、同输入同输出。
 * 依赖     : 无 DL_ 内部依赖（本批自足实现）
 * 修订历史 :
 *        2026-11-23  v1.0.0  R78-B1 对齐取整族模板派生首版
 *        2026-11-24  v1.0.1  R79-F1 修 DINT 回绕（R78 闸 L1 阻断项）：
 *                    ① 进位侧 nLo + nMultiple 在 nLo 接近 DINT_MAX 时溢出回绕成负数
 *                       （例：nValue=DINT_MAX-1, nMultiple=4 → 结果变负）；
 *                    ② 退位侧 nLo - nMultiple 在 nLo 接近 DINT_MIN 时同理溢出。
 *                    修法：加显式上/下饱和闸 —— 进位前判 nLo > DINT_MAX - nMultiple，
 *                    退位前判 nLo < DINT_MIN + nMultiple，命中即钳到域端点并置
 *                    bSat := TRUE（饱和出口），不再做算术进位 / 退位。
 *                    该闸使"整数域内不可表示的四舍五入结果"饱和而非回绕，符合安全侧
 *                    优先（宁可饱和到端点让上位机看见 bSat，不可回绕成反向大数）。
 * 红线自检 : R1 零全局 R2 零%I/%Q R3 纯IEC R4 非法倍数返 0 + 比较用 nHalf
 *            避免 nRem*2 溢出 + 上/下饱和闸防 nLo±nMultiple 回绕 (v1.0.1)
 *            R5 双语注释 R6 N/A（无状态机） R7 N/A R10 无构造式转换
 *============================================================================*)
FUNCTION FC_DL_RoundToMultipleInt : DINT
VAR_INPUT
    nValue : DINT;          // 输入整数 / Input integer value
    nMultiple : DINT;       // 对齐倍数，须 > 0 / Alignment multiple, must be > 0
END_VAR
VAR_OUTPUT
    bSat : BOOL;            // 结果已饱和到 DINT 域端点（未真四舍五入）/ Result saturated at the DINT domain end
    bError : BOOL;          // 倍数非法（<= 0）/ Invalid multiple (<= 0)
END_VAR
VAR
    nLo : DINT;             // 向零截断的基准倍数值 / Truncated-toward-zero base multiple
    nRem : DINT;            // 余量，符号随被除数，绝对值 < nMultiple / Remainder, |nRem| < nMultiple
    nHalf : DINT;           // 倍数半值（向下取整） / Floor half of the multiple
END_VAR
VAR CONSTANT
    DL_RMI_MAX : DINT := 2147483647;    // DINT 上端 / Upper end of DINT
    DL_RMI_MIN : DINT := -2147483648;   // DINT 下端 / Lower end of DINT
END_VAR
bSat := FALSE;                          // 饱和标志每调用先清 / Clear the saturation flag every call
bError := FALSE;                        // 错误标志每调用先清 / Clear the error flag every call
IF nMultiple <= 0 THEN
    bError := TRUE;                     // 倍数非法回执 / Invalid multiple receipt
    FC_DL_RoundToMultipleInt := 0;      // 非法倍数返 0 / Invalid multiple returns 0
    RETURN;
END_IF
nLo := (nValue / nMultiple) * nMultiple;    // 整除截取得基准 / Base via integer division truncation
nRem := nValue - nLo;                       // 余量 / Remainder in (-nMultiple, nMultiple)
nHalf := nMultiple / 2;                     // 半值基准，免 nRem*2 溢出 / Half reference avoids nRem*2 overflow
IF nRem >= 0 THEN
    IF (nRem > nHalf) OR ((nRem = nHalf) AND ((nMultiple MOD 2) = 0)) THEN
        IF nLo > (DL_RMI_MAX - nMultiple) THEN
            nLo := DL_RMI_MAX;              // 进位将溢出 → 饱和到上端 / Round up would overflow, saturate high
            bSat := TRUE;                   // 置饱和标志 / Raise the saturation flag
        ELSE
            nLo := nLo + nMultiple;         // 正余量过半进位 / Round up at half
        END_IF
    END_IF
ELSIF (-nRem > nHalf) OR ((-nRem = nHalf) AND ((nMultiple MOD 2) = 0)) THEN
    IF nLo < (DL_RMI_MIN + nMultiple) THEN
        nLo := DL_RMI_MIN;                  // 退位将溢出 → 饱和到下端 / Round down would overflow, saturate low
        bSat := TRUE;                       // 置饱和标志 / Raise the saturation flag
    ELSE
        nLo := nLo - nMultiple;             // 负余量过半退位 / Round down at half
    END_IF
END_IF
FC_DL_RoundToMultipleInt := nLo;            // 输出四舍五入结果 / Output rounded result
END_FUNCTION

(* ---- FC_DL_RoundToMultipleReal.st ---- *)
(*==============================================================================
 * 组件名称 : FC_DL_RoundToMultipleReal ｜ 子库 : DL_MathData ｜ v1.0.0 ｜ 2026-11-23
 * 平台     : CODESYS 3.5 / TwinCAT 3 / InoProShop / Machine Expert（纯 IEC，无厂商库）
 * 功能简介 : 实数四舍五入到 fMultiple 的最近倍数。先除到倍数域，经标准
 *            就近舍入型转换 REAL_TO_DINT 取最近整倍数序号，再映射回倍数域。
 * 契约     : 返回四舍五入后的倍数值 [fMultiple 单位]；fMultiple <= 0 或
 *            输入 NaN/Inf 恒返回 0.0；商超出 DINT 安全域时按原值近直返；
 *            纯函数无状态、同输入同输出。
 * 依赖     : 无 DL_ 内部依赖（本批自足实现）
 * 红线自检 : R1 零全局 R2 零%I/%Q R3 纯IEC（*_TO_* 显式转换）R4 非法倍数/
 *            NaN/Inf 返 0 + 商域闸防 REAL_TO_DINT 溢出 R5 双语注释
 *            R6 N/A（无状态机） R7 N/A（无定时器实例）
 * 修订历史 : 2026-11-23 R78-B1 对齐取整族模板派生首版
 *============================================================================*)
FUNCTION FC_DL_RoundToMultipleReal : REAL
VAR_INPUT
    fValue : REAL;          // 输入实数 / Input real value
    fMultiple : REAL;       // 对齐倍数，须 > 0 / Multiple, must be > 0
END_VAR
VAR
    fQ : REAL;              // 倍数域商 / Ratio in multiple domain
    nQ : DINT;              // 最近整倍数序号 / Nearest multiple index
END_VAR
VAR CONSTANT
    DL_Q_SAFE_MAX : REAL := 2.0E9;      // DINT 安全商上限，防转换溢出 / Safe ratio cap guarding conversion overflow
END_VAR
IF (fMultiple <= 0.0) OR (fValue <> fValue) OR ((fValue - fValue) <> 0.0) THEN
    FC_DL_RoundToMultipleReal := 0.0;   // 非法倍数或 NaN/Inf 输入返 0 / Invalid multiple or NaN/Inf returns 0
    RETURN;
END_IF
fQ := fValue / fMultiple;                           // 商 / Ratio
IF (fQ <> fQ) OR ((fQ - fQ) <> 0.0) OR (fQ > DL_Q_SAFE_MAX) OR (fQ < -DL_Q_SAFE_MAX) THEN
    FC_DL_RoundToMultipleReal := fQ * fMultiple;    // 商 NaN/Inf/超域按原值近直返 / NaN/Inf/out-of-domain ratio returns near-original
    RETURN;
END_IF
nQ := REAL_TO_DINT(fQ);                             // 最近邻取整（IEC 实转整为就近舍入）/ Round to nearest via typed conversion
FC_DL_RoundToMultipleReal := DINT_TO_REAL(nQ) * fMultiple;      // 映射回倍数域 / Map back to multiple domain
END_FUNCTION

(* ---- FC_DL_SatAddDint.st ---- *)
(*
  FC_DL_SatAddDint —— DINT 加法饱和，上下界检测
  分类：DL_MathData | 复杂度：2 | 轮次：R86
  开源溯源：道莅原创（clean-room 自研，纯 IEC 61131-3 通用算法），无外部代码引用
  许可证：MIT
  职责：有符号双整数加法，越界时钳到 DINT 上下界并置 xSat；用「带符号双侧直比」判溢出，
        禁用 ABS 单侧比较（ABS(DINT_MIN) 自身会溢出）。
  契约：diA / diB 加数；diOut 饱和和；xSat 报告饱和（信息级）。DINT 上下界在本文件内定义，不跨文件引用。
  边界：① 同号才可能溢出，异号必不溢出；② 上界判据 diA > MAX - diB（diB > 0），下界判 diA < MIN - diB（diB < 0）；
        ③ 零全局、零物理地址、零库件依赖。
*)
FUNCTION FC_DL_SatAddDint : DINT
VAR_INPUT
    diA : DINT := 0;                  // 加数 A [—] / The addend A
    diB : DINT := 0;                  // 加数 B [—] / The addend B
END_VAR
VAR_OUTPUT
    xSat : BOOL;                      // 饱和发生标志（信息级） [—] / The saturation flag, informational
END_VAR
VAR CONSTANT
    DL_DINT_MAX : DINT := 2147483647; // DINT 上界（本件私有） [-] / The DINT maximum, private to this file
    DL_DINT_MIN : DINT := -2147483647 - 1; // DINT 下界（本件私有，减法写法避免字面量越域） [-] / The DINT minimum
END_VAR

xSat := FALSE;                                        // 饱和标志预置假 / preset the saturation flag false
IF (diB > 0) AND (diA > (DL_DINT_MAX - diB)) THEN     // 正加数上溢判据（双侧直比） / the positive overflow test
    FC_DL_SatAddDint := DL_DINT_MAX;                  // 钳到上界 / clamp to the maximum
    xSat := TRUE;                                     // 置饱和标志 / raise the saturation flag
ELSIF (diB < 0) AND (diA < (DL_DINT_MIN - diB)) THEN  // 负加数下溢判据（双侧直比） / the negative overflow test
    FC_DL_SatAddDint := DL_DINT_MIN;                  // 钳到下界 / clamp to the minimum
    xSat := TRUE;                                     // 置饱和标志 / raise the saturation flag
ELSE
    FC_DL_SatAddDint := diA + diB;                    // 界内直接相加 / the safe addition
END_IF
END_FUNCTION

(* ---- FC_DL_SatAddLreal.st ---- *)
(*
  FC_DL_SatAddLreal —— LREAL 加法饱和加非有限值闸
  分类：DL_MathData | 复杂度：2 | 轮次：R86
  开源溯源：道莅原创（clean-room 自研，纯 IEC 61131-3 通用算法），无外部代码引用
  许可证：MIT
  职责：实数加法后按 [fMin, fMax] 饱和；四个浮点入参逐一做非有限闸（NaN 自反判、Inf 用 1.0E30 绝对上限判），
        任一非法即 fOut 归零并置 xValid = FALSE。
  契约：fA / fB 加数、fMin / fMax 饱和区间；fOut 结果；xSat 报告饱和；xValid 结果可信。
  边界：① 区间倒置判非法；② 求和结果再做一次非有限自检（Inf 求和路径）；
        ③ 零全局、零物理地址、零库件依赖。
*)
FUNCTION FC_DL_SatAddLreal : LREAL
VAR_INPUT
    fA   : LREAL := 0.0;              // 加数 A [工程单位] / The addend A
    fB   : LREAL := 0.0;              // 加数 B [工程单位] / The addend B
    fMin : LREAL := -1000.0;          // 饱和下限 [工程单位] / The saturation low limit
    fMax : LREAL := 1000.0;           // 饱和上限 [工程单位] / The saturation high limit
END_VAR
VAR_OUTPUT
    xSat   : BOOL;                    // 饱和发生标志（信息级） [—] / The saturation flag, informational
    xValid : BOOL;                    // 结果可信 [—] / The result is valid
END_VAR
VAR
    fSum : LREAL;                     // 求和中间量 [工程单位] / The sum intermediate
END_VAR
VAR CONSTANT
    DL_AL_INF : LREAL := 1.0E30;      // 非有限 / 越界判据上限 [-] / The magnitude gate
    DL_AL_Z   : LREAL := 0.0;         // 浮点零常量 [工程单位] / The floating point zero constant
END_VAR

xSat := FALSE;                                        // 饱和标志预置假 / preset the saturation flag false
xValid := FALSE;                                      // 可信位预置假 / preset the valid flag false
FC_DL_SatAddLreal := DL_AL_Z;                         // 返回值预置零 / preset the return zero
IF (fA <> fA) OR (ABS(fA) > DL_AL_INF) THEN           // 加数 A 非有限闸 / the addend A gate
    FC_DL_SatAddLreal := DL_AL_Z;                     // 非有限归零 / zero the non finite input
ELSIF (fB <> fB) OR (ABS(fB) > DL_AL_INF) THEN        // 加数 B 非有限闸 / the addend B gate
    FC_DL_SatAddLreal := DL_AL_Z;                     // 非有限归零 / zero the non finite input
ELSIF (fMin <> fMin) OR (ABS(fMin) > DL_AL_INF) THEN  // 下限非有限闸 / the low limit gate
    FC_DL_SatAddLreal := DL_AL_Z;                     // 非有限归零 / zero the non finite input
ELSIF (fMax <> fMax) OR (ABS(fMax) > DL_AL_INF) THEN  // 上限非有限闸 / the high limit gate
    FC_DL_SatAddLreal := DL_AL_Z;                     // 非有限归零 / zero the non finite input
ELSIF fMax < fMin THEN                                // 饱和区间倒置 / the saturated band is inverted
    FC_DL_SatAddLreal := DL_AL_Z;                     // 非法区间归零 / zero on an invalid band
ELSE
    fSum := fA + fB;                                  // 求和 [工程单位] / the sum
    IF fSum <> fSum THEN                              // 求和结果非有限自检 / the sum self check
        FC_DL_SatAddLreal := DL_AL_Z;                 // 非有限归零 / zero the non finite sum
    ELSIF fSum > fMax THEN                            // 上越界 / above the high limit
        FC_DL_SatAddLreal := fMax;                    // 钳到上限 [工程单位] / clamp to the high limit
        xSat := TRUE;                                 // 置饱和标志 / raise the saturation flag
        xValid := TRUE;                               // 饱和输出仍可信 / a saturated output is still valid
    ELSIF fSum < fMin THEN                            // 下越界 / below the low limit
        FC_DL_SatAddLreal := fMin;                    // 钳到下限 [工程单位] / clamp to the low limit
        xSat := TRUE;                                 // 置饱和标志 / raise the saturation flag
        xValid := TRUE;                               // 饱和输出仍可信 / a saturated output is still valid
    ELSE
        FC_DL_SatAddLreal := fSum;                    // 界内直接输出 / the in range sum
        xValid := TRUE;                               // 结果可信 / the result is valid
    END_IF
END_IF
END_FUNCTION

(* ---- FC_DL_SatClampLrealBand.st ---- *)
(*
  FC_DL_SatClampLrealBand —— LREAL 区间钳位，带上下限合法性自检
  分类：DL_MathData | 复杂度：1 | 轮次：R86
  开源溯源：道莅原创（clean-room 自研，纯 IEC 61131-3 通用算法），无外部代码引用
  许可证：MIT
  职责：把输入钳到 [fMin, fMax]；钳位前先自检区间合法性（fMax 必须 >= fMin）与三个浮点入参的非有限性，
        任一非法即 fOut 给下限哨兵并置 xValid = FALSE。
  契约：fIn 输入、fMin / fMax 钳位区间；fOut 钳位结果；xClamped 报告发生钳位；xValid 结果可信。
  边界：① 区间倒置判非法（不静默交换，交换会掩盖上游配置错误）；② 三个浮点入参逐一非有限闸；
        ③ 零全局、零物理地址、零库件依赖。
*)
FUNCTION FC_DL_SatClampLrealBand : LREAL
VAR_INPUT
    fIn  : LREAL := 0.0;              // 输入值 [工程单位] / The input value
    fMin : LREAL := -1000.0;          // 钳位下限 [工程单位] / The clamp low limit
    fMax : LREAL := 1000.0;           // 钳位上限 [工程单位] / The clamp high limit
END_VAR
VAR_OUTPUT
    xClamped : BOOL;                  // 发生钳位（信息级） [—] / A clamp occurred, informational
    xValid   : BOOL;                  // 区间与输入合法 [—] / The band and the input are valid
END_VAR
VAR CONSTANT
    DL_CL_INF : LREAL := 1.0E30;      // 非有限 / 越界判据上限 [-] / The magnitude gate
    DL_CL_Z   : LREAL := 0.0;         // 浮点零常量 [工程单位] / The floating point zero constant
END_VAR

xClamped := FALSE;                                    // 钳位标志预置假 / preset the clamp flag false
xValid := FALSE;                                      // 可信位预置假 / preset the valid flag false
FC_DL_SatClampLrealBand := DL_CL_Z;                   // 返回值预置零 / preset the return zero
IF (fIn <> fIn) OR (ABS(fIn) > DL_CL_INF) THEN        // 输入非有限闸 / the input gate
    FC_DL_SatClampLrealBand := fMin;                  // 非有限输入给下限哨兵 / the low limit sentinel
ELSIF (fMin <> fMin) OR (ABS(fMin) > DL_CL_INF) THEN  // 下限非有限闸 / the low limit gate
    FC_DL_SatClampLrealBand := DL_CL_Z;               // 下限非法归零 / zero on an invalid limit
ELSIF (fMax <> fMax) OR (ABS(fMax) > DL_CL_INF) THEN  // 上限非有限闸 / the high limit gate
    FC_DL_SatClampLrealBand := DL_CL_Z;               // 上限非法归零 / zero on an invalid limit
ELSIF fMax < fMin THEN                                // 区间倒置（配置错误的显式拒绝） / the inverted band
    FC_DL_SatClampLrealBand := fMin;                  // 倒置区间给下限哨兵 / the low limit sentinel
ELSE
    IF fIn > fMax THEN                                // 上越界钳位 / clamp the high side
        FC_DL_SatClampLrealBand := fMax;              // 钳到上限 [工程单位] / clamp to the high limit
        xClamped := TRUE;                             // 置钳位标志 / raise the clamp flag
    ELSIF fIn < fMin THEN                             // 下越界钳位 / clamp the low side
        FC_DL_SatClampLrealBand := fMin;              // 钳到下限 [工程单位] / clamp to the low limit
        xClamped := TRUE;                             // 置钳位标志 / raise the clamp flag
    ELSE
        FC_DL_SatClampLrealBand := fIn;               // 界内直接输出 [工程单位] / the in range value
    END_IF
    xValid := TRUE;                                   // 区间与输入合法 / the band and the input are valid
END_IF
END_FUNCTION

(* ---- FC_DL_SatMulDint.st ---- *)
(*
  FC_DL_SatMulDint —— DINT 乘法饱和，先判溢出条件再乘
  分类：DL_MathData | 复杂度：2 | 轮次：R86
  开源溯源：道莅原创（clean-room 自研，纯 IEC 61131-3 通用算法），无外部代码引用
  许可证：MIT
  职责：有符号双整数乘法，先做「除后比较」溢出判定再执行乘法，越界钳到 DINT 上下界并置 xSat。
  契约：diA / diB 乘数；diOut 饱和积；xSat 报告饱和（信息级）。DINT 上下界在本文件内定义。
  边界：① 零乘数先短路；② DINT_MIN 单独分支（ABS(DINT_MIN) 会溢出，禁走 ABS 路径）；
        ③ 一般情形用 |a| > MAX / |b| 的整除判据（整除结果偏保守，安全方向）；
        ④ 零全局、零物理地址、零库件依赖。
*)
FUNCTION FC_DL_SatMulDint : DINT
VAR_INPUT
    diA : DINT := 0;                  // 乘数 A [—] / The multiplier A
    diB : DINT := 0;                  // 乘数 B [—] / The multiplier B
END_VAR
VAR_OUTPUT
    xSat : BOOL;                      // 饱和发生标志（信息级） [—] / The saturation flag, informational
END_VAR
VAR
    xNeg : BOOL;                      // 积的符号（异号） [—] / The product sign, true when opposite
END_VAR
VAR CONSTANT
    DL_DINT_MAX : DINT := 2147483647; // DINT 上界（本件私有） [-] / The DINT maximum, private to this file
    DL_DINT_MIN : DINT := -2147483647 - 1; // DINT 下界（本件私有） [-] / The DINT minimum, private to this file
END_VAR

xSat := FALSE;                                        // 饱和标志预置假 / preset the saturation flag false
xNeg := ((diA > 0) AND (diB < 0)) OR ((diA < 0) AND (diB > 0)); // 异号判定 / the opposite sign test
IF (diA = 0) OR (diB = 0) THEN                        // 零乘数短路（不溢出） / a zero multiplier never overflows
    FC_DL_SatMulDint := 0;                            // 积为零 / the product is zero
ELSIF diB = 1 THEN                                    // 乘一保持原值 / multiply by one keeps the value
    FC_DL_SatMulDint := diA;                          // 返回被乘数 / return the other operand
ELSIF diA = 1 THEN                                    // 乘一保持原值 / multiply by one keeps the value
    FC_DL_SatMulDint := diB;                          // 返回被乘数 / return the other operand
ELSIF diB = -1 THEN                                   // 乘负一（DINT_MIN 例外） / multiply by minus one
    IF diA = DL_DINT_MIN THEN                         // 唯一上溢组合 / the only overflowing combination
        FC_DL_SatMulDint := DL_DINT_MAX;              // 钳到上界 / clamp to the maximum
        xSat := TRUE;                                 // 置饱和标志 / raise the saturation flag
    ELSE
        FC_DL_SatMulDint := 0 - diA;                  // 取负（界内） / the in range negation
    END_IF
ELSIF diA = -1 THEN                                   // 乘负一（DINT_MIN 例外） / multiply by minus one
    IF diB = DL_DINT_MIN THEN                         // 唯一上溢组合 / the only overflowing combination
        FC_DL_SatMulDint := DL_DINT_MAX;              // 钳到上界 / clamp to the maximum
        xSat := TRUE;                                 // 置饱和标志 / raise the saturation flag
    ELSE
        FC_DL_SatMulDint := 0 - diB;                  // 取负（界内） / the in range negation
    END_IF
ELSIF (diA = DL_DINT_MAX) OR (diB = DL_DINT_MAX) OR (diA = DL_DINT_MIN) OR (diB = DL_DINT_MIN) THEN
    IF xNeg THEN                                      // 异号，积为负，溢出下界 / opposite signs underflow
        FC_DL_SatMulDint := DL_DINT_MIN;              // 钳到下界 / clamp to the minimum
    ELSE                                              // 同号，积为正，溢出上界 / the same signs overflow high
        FC_DL_SatMulDint := DL_DINT_MAX;              // 钳到上界 / clamp to the maximum
    END_IF
    xSat := TRUE;                                     // 置饱和标志 / raise the saturation flag
ELSIF ABS(diA) > (DL_DINT_MAX / ABS(diB)) THEN        // 除后比较（两乘数均已排除 DINT_MIN，ABS 安全） / the divide test
    IF xNeg THEN                                      // 异号下溢 / the negative overflow
        FC_DL_SatMulDint := DL_DINT_MIN;              // 钳到下界 / clamp to the minimum
    ELSE                                              // 同号上溢 / the positive overflow
        FC_DL_SatMulDint := DL_DINT_MAX;              // 钳到上界 / clamp to the maximum
    END_IF
    xSat := TRUE;                                     // 置饱和标志 / raise the saturation flag
ELSE
    FC_DL_SatMulDint := diA * diB;                    // 界内直接相乘 / the safe multiplication
END_IF
END_FUNCTION

(* ---- FC_DL_SatMulLreal.st ---- *)
(*
  FC_DL_SatMulLreal —— LREAL 乘法饱和加非有限值闸
  分类：DL_MathData | 复杂度：2 | 轮次：R86
  开源溯源：道莅原创（clean-room 自研，纯 IEC 61131-3 通用算法），无外部代码引用
  许可证：MIT
  职责：实数乘法后按 [fMin, fMax] 饱和；四个浮点入参逐一非有限闸，任一非法即归零并置 xValid = FALSE。
  契约：fA / fB 乘数、fMin / fMax 饱和区间；fOut 结果；xSat 报告饱和；xValid 结果可信。
  边界：① 区间倒置判非法；② 乘积非有限自检（1.0E30 量级输入相乘可达 1.0E60，仍属有限，但保留自检闸）；
        ③ 零乘数短路为 0（不进入饱和路径）；④ 零全局、零物理地址、零库件依赖。
*)
FUNCTION FC_DL_SatMulLreal : LREAL
VAR_INPUT
    fA   : LREAL := 1.0;              // 乘数 A [工程单位] / The multiplier A
    fB   : LREAL := 1.0;              // 乘数 B [—] / The multiplier B
    fMin : LREAL := -1000.0;          // 饱和下限 [工程单位] / The saturation low limit
    fMax : LREAL := 1000.0;           // 饱和上限 [工程单位] / The saturation high limit
END_VAR
VAR_OUTPUT
    xSat   : BOOL;                    // 饱和发生标志（信息级） [—] / The saturation flag, informational
    xValid : BOOL;                    // 结果可信 [—] / The result is valid
END_VAR
VAR
    fProd : LREAL;                    // 乘积中间量 [工程单位] / The product intermediate
END_VAR
VAR CONSTANT
    DL_ML_INF : LREAL := 1.0E30;      // 非有限 / 越界判据上限 [-] / The magnitude gate
    DL_ML_Z   : LREAL := 0.0;         // 浮点零常量 [工程单位] / The floating point zero constant
END_VAR

xSat := FALSE;                                        // 饱和标志预置假 / preset the saturation flag false
xValid := FALSE;                                      // 可信位预置假 / preset the valid flag false
FC_DL_SatMulLreal := DL_ML_Z;                         // 返回值预置零 / preset the return zero
IF (fA <> fA) OR (ABS(fA) > DL_ML_INF) THEN           // 乘数 A 非有限闸 / the multiplier A gate
    FC_DL_SatMulLreal := DL_ML_Z;                     // 非有限归零 / zero the non finite input
ELSIF (fB <> fB) OR (ABS(fB) > DL_ML_INF) THEN        // 乘数 B 非有限闸 / the multiplier B gate
    FC_DL_SatMulLreal := DL_ML_Z;                     // 非有限归零 / zero the non finite input
ELSIF (fMin <> fMin) OR (ABS(fMin) > DL_ML_INF) THEN  // 下限非有限闸 / the low limit gate
    FC_DL_SatMulLreal := DL_ML_Z;                     // 非有限归零 / zero the non finite input
ELSIF (fMax <> fMax) OR (ABS(fMax) > DL_ML_INF) THEN  // 上限非有限闸 / the high limit gate
    FC_DL_SatMulLreal := DL_ML_Z;                     // 非有限归零 / zero the non finite input
ELSIF fMax < fMin THEN                                // 饱和区间倒置 / the saturated band is inverted
    FC_DL_SatMulLreal := DL_ML_Z;                     // 非法区间归零 / zero on an invalid band
ELSE
    fProd := fA * fB;                                 // 求积 [工程单位] / the product
    IF fProd <> fProd THEN                            // 乘积非有限自检 / the product self check
        FC_DL_SatMulLreal := DL_ML_Z;                 // 非有限归零 / zero the non finite product
    ELSIF fProd > fMax THEN                           // 上越界 / above the high limit
        FC_DL_SatMulLreal := fMax;                    // 钳到上限 [工程单位] / clamp to the high limit
        xSat := TRUE;                                 // 置饱和标志 / raise the saturation flag
        xValid := TRUE;                               // 饱和输出仍可信 / a saturated output is still valid
    ELSIF fProd < fMin THEN                           // 下越界 / below the low limit
        FC_DL_SatMulLreal := fMin;                    // 钳到下限 [工程单位] / clamp to the low limit
        xSat := TRUE;                                 // 置饱和标志 / raise the saturation flag
        xValid := TRUE;                               // 饱和输出仍可信 / a saturated output is still valid
    ELSE
        FC_DL_SatMulLreal := fProd;                   // 界内直接输出 / the in range product
        xValid := TRUE;                               // 结果可信 / the result is valid
    END_IF
END_IF
END_FUNCTION

(* ---- FC_DL_SatNegDint.st ---- *)
(*
  FC_DL_SatNegDint —— DINT 取负饱和，DINT_MIN 不回绕
  分类：DL_MathData | 复杂度：1 | 轮次：R86
  开源溯源：道莅原创（clean-room 自研，纯 IEC 61131-3 通用算法），无外部代码引用
  许可证：MIT
  职责：双整数取负；DINT_MIN 的相反数超出 DINT 上界，饱和到 DINT_MAX 并置 xSat，绝不回绕成负数。
  契约：diIn 输入；diOut 结果；xSat 报告边界饱和（信息级）。DINT 上下界在本文件内定义。
  边界：不使用一元负号直接作用于 DINT（DINT_MIN 回绕），改用 0 - diIn 并前置边界分支；
        零全局、零物理地址、零库件依赖。
*)
FUNCTION FC_DL_SatNegDint : DINT
VAR_INPUT
    diIn : DINT := 0;                 // 输入操作数 [—] / The input operand
END_VAR
VAR_OUTPUT
    xSat : BOOL;                      // 边界饱和标志（信息级） [—] / The boundary saturation flag
END_VAR
VAR CONSTANT
    DL_DINT_MAX : DINT := 2147483647; // DINT 上界（本件私有） [-] / The DINT maximum, private to this file
    DL_DINT_MIN : DINT := -2147483647 - 1; // DINT 下界（本件私有） [-] / The DINT minimum, private to this file
END_VAR

xSat := FALSE;                                        // 饱和标志预置假 / preset the saturation flag false
IF diIn = DL_DINT_MIN THEN                            // 唯一回绕点 / the only wrapping input
    FC_DL_SatNegDint := DL_DINT_MAX;                  // 饱和到上界 / saturate to the maximum
    xSat := TRUE;                                     // 置饱和标志 / raise the saturation flag
ELSE
    FC_DL_SatNegDint := 0 - diIn;                     // 双字域取负（界内安全） / the in range negation
END_IF
END_FUNCTION

(* ---- FC_DL_SatScaleLreal.st ---- *)
(*
  FC_DL_SatScaleLreal —— LREAL 增益缩放饱和
  分类：DL_MathData | 复杂度：2 | 轮次：R86
  开源溯源：道莅原创（clean-room 自研，纯 IEC 61131-3 通用算法），无外部代码引用
  许可证：MIT
  职责：实数增益缩放（out = fIn * fGain）后按 [fMin, fMax] 饱和；四个浮点入参逐一非有限闸，
        任一非法即归零并置 xValid = FALSE。
  契约：fIn 输入、fGain 增益、fMin / fMax 饱和区间；fOut 结果；xSat 报告饱和；xValid 结果可信。
  边界：① 区间倒置判非法；② 乘积非有限自检；③ 增益为 0 时输出 0（不进入饱和路径）；
        ④ 零全局、零物理地址、零库件依赖。
*)
FUNCTION FC_DL_SatScaleLreal : LREAL
VAR_INPUT
    fIn   : LREAL := 0.0;             // 输入值 [工程单位] / The input value
    fGain : LREAL := 1.0;             // 缩放增益 [—] / The scaling gain
    fMin  : LREAL := -1000.0;         // 饱和下限 [工程单位] / The saturation low limit
    fMax  : LREAL := 1000.0;          // 饱和上限 [工程单位] / The saturation high limit
END_VAR
VAR_OUTPUT
    xSat   : BOOL;                    // 饱和发生标志（信息级） [—] / The saturation flag, informational
    xValid : BOOL;                    // 结果可信 [—] / The result is valid
END_VAR
VAR
    fScaled : LREAL;                  // 缩放中间量 [工程单位] / The scaled intermediate
END_VAR
VAR CONSTANT
    DL_SL_INF : LREAL := 1.0E30;      // 非有限 / 越界判据上限 [-] / The magnitude gate
    DL_SL_Z   : LREAL := 0.0;         // 浮点零常量 [工程单位] / The floating point zero constant
END_VAR

xSat := FALSE;                                        // 饱和标志预置假 / preset the saturation flag false
xValid := FALSE;                                      // 可信位预置假 / preset the valid flag false
FC_DL_SatScaleLreal := DL_SL_Z;                       // 返回值预置零 / preset the return zero
IF (fIn <> fIn) OR (ABS(fIn) > DL_SL_INF) THEN        // 输入非有限闸 / the input gate
    FC_DL_SatScaleLreal := DL_SL_Z;                   // 非有限归零 / zero the non finite input
ELSIF (fGain <> fGain) OR (ABS(fGain) > DL_SL_INF) THEN // 增益非有限闸 / the gain gate
    FC_DL_SatScaleLreal := DL_SL_Z;                   // 非有限归零 / zero the non finite gain
ELSIF (fMin <> fMin) OR (ABS(fMin) > DL_SL_INF) THEN  // 下限非有限闸 / the low limit gate
    FC_DL_SatScaleLreal := DL_SL_Z;                   // 非有限归零 / zero the non finite limit
ELSIF (fMax <> fMax) OR (ABS(fMax) > DL_SL_INF) THEN  // 上限非有限闸 / the high limit gate
    FC_DL_SatScaleLreal := DL_SL_Z;                   // 非有限归零 / zero the non finite limit
ELSIF fMax < fMin THEN                                // 饱和区间倒置 / the saturated band is inverted
    FC_DL_SatScaleLreal := DL_SL_Z;                   // 非法区间归零 / zero on an invalid band
ELSE
    fScaled := fIn * fGain;                           // 增益缩放 [工程单位] / the scaled value
    IF fScaled <> fScaled THEN                        // 缩放结果非有限自检 / the scaled value self check
        FC_DL_SatScaleLreal := DL_SL_Z;               // 非有限归零 / zero the non finite value
    ELSIF fScaled > fMax THEN                         // 上越界 / above the high limit
        FC_DL_SatScaleLreal := fMax;                  // 钳到上限 [工程单位] / clamp to the high limit
        xSat := TRUE;                                 // 置饱和标志 / raise the saturation flag
        xValid := TRUE;                               // 饱和输出仍可信 / a saturated output is still valid
    ELSIF fScaled < fMin THEN                         // 下越界 / below the low limit
        FC_DL_SatScaleLreal := fMin;                  // 钳到下限 [工程单位] / clamp to the low limit
        xSat := TRUE;                                 // 置饱和标志 / raise the saturation flag
        xValid := TRUE;                               // 饱和输出仍可信 / a saturated output is still valid
    ELSE
        FC_DL_SatScaleLreal := fScaled;               // 界内直接输出 / the in range value
        xValid := TRUE;                               // 结果可信 / the result is valid
    END_IF
END_IF
END_FUNCTION

(* ---- FC_DL_SatSumArrayDint.st ---- *)
(*
  FC_DL_SatSumArrayDint —— DINT 定长数组累加饱和，逐项防溢出
  分类：DL_MathData | 复杂度：2 | 轮次：R86
  开源溯源：道莅原创（clean-room 自研，纯 IEC 61131-3 通用算法），无外部代码引用
  许可证：MIT
  职责：对定长 8 元 DINT 数组的前 nCnt 项求和，每加一项前做「双侧直比」溢出判定，
        一旦越界即钳到 DINT 上下界、置 xSat 并停止累加（饱和语义，不做回绕）。
  契约：arrIn 输入数组（显式定长，R15）、nCnt 参与项数（0..8，越界自动截断）；diOut 饱和和；
        nUsed 实际参与项数；xSat 报告饱和。DINT 上下界在本文件内定义。
  边界：① 项数越域截断到 0..8；② 逐项溢出前置判定（禁 ABS 单侧比较）；③ 饱和即终止，结果单调可信；
        ④ 零全局、零物理地址、零库件依赖。
*)
FUNCTION FC_DL_SatSumArrayDint : DINT
VAR_INPUT
    arrIn : ARRAY[0..7] OF DINT;      // 输入数组（显式定长 8 元） [—] / The fixed length input array
    nCnt  : INT := 8;                 // 参与累加的项数（0..8） [个] / The number of items to sum
END_VAR
VAR_OUTPUT
    nUsed : INT;                      // 实际参与累加的项数 [个] / The number of items actually summed
    xSat  : BOOL;                     // 饱和发生标志（信息级） [—] / The saturation flag, informational
END_VAR
VAR
    i     : INT;                      // 遍历索引 [下标] / The traversal index
    diAcc : DINT;                     // 累加器 [—] / The accumulator
    diItem : DINT;                    // 当前项 [—] / The current item
    xStop : BOOL;                     // 饱和终止标志 [—] / The saturation stop flag
END_VAR
VAR CONSTANT
    DL_DINT_MAX : DINT := 2147483647; // DINT 上界（本件私有） [-] / The DINT maximum, private to this file
    DL_DINT_MIN : DINT := -2147483647 - 1; // DINT 下界（本件私有） [-] / The DINT minimum, private to this file
    DL_SA_NMAX  : INT := 8;           // 数组容量 [个] / The array capacity
    DL_SA_Z     : INT := 0;           // 整型零常量 [个] / The integer zero constant
END_VAR

FC_DL_SatSumArrayDint := 0;                           // 返回值预置零 / preset the return zero
xSat := FALSE;                                        // 饱和标志预置假 / preset the saturation flag false
nUsed := DL_SA_Z;                                     // 参与项数预置零 [个] / preset the used count zero
diAcc := 0;                                           // 累加器清零 [—] / clear the accumulator
xStop := FALSE;                                       // 终止标志预置假 / preset the stop flag false
IF nCnt < DL_SA_Z THEN                                // 项数下越界 / the count below the domain
    nCnt := DL_SA_Z;                                  // 截断到零 [个] / truncate to zero
END_IF
IF nCnt > DL_SA_NMAX THEN                             // 项数上越界 / the count above the capacity
    nCnt := DL_SA_NMAX;                               // 截断到容量 [个] / truncate to the capacity
END_IF
i := DL_SA_Z;                                         // 索引从零起 / start from the first item
WHILE (i < nCnt) AND NOT xStop DO                     // 显式递增逐项累加 / accumulate item by item
    diItem := arrIn[i];                               // 取当前项 [—] / take the current item
    IF (diItem > 0) AND (diAcc > (DL_DINT_MAX - diItem)) THEN // 正项上溢前置判定 / the positive overflow test
        diAcc := DL_DINT_MAX;                         // 钳到上界 / clamp to the maximum
        xSat := TRUE;                                 // 置饱和标志 / raise the saturation flag
        xStop := TRUE;                                // 终止后续累加 / stop the accumulation
    ELSIF (diItem < 0) AND (diAcc < (DL_DINT_MIN - diItem)) THEN // 负项下溢前置判定 / the negative overflow test
        diAcc := DL_DINT_MIN;                         // 钳到下界 / clamp to the minimum
        xSat := TRUE;                                 // 置饱和标志 / raise the saturation flag
        xStop := TRUE;                                // 终止后续累加 / stop the accumulation
    ELSE
        diAcc := diAcc + diItem;                      // 界内累加 / the safe accumulation
        nUsed := nUsed + 1;                           // 计入参与项数 [个] / count the summed item
    END_IF
    i := i + 1;                                       // 索引递增 [下标] / increment the index
END_WHILE
FC_DL_SatSumArrayDint := diAcc;                       // 饱和和出口 [—] / publish the saturated sum
END_FUNCTION

(* ---- FC_DL_SaturateDecr.st ---- *)
(*==============================================================================
 * 组件名称 (Component)  : FC_DL_SaturateDecr
 * 所属子库 (Sublibrary) : DL_MathData ｜ 版本 (Version) : 1.0.0 ｜ 2026-11-23
 * 兼容性   (Platform)   : CODESYS 3.5+ / TwinCAT 3 / 汇川 InoProShop / 施耐德 Machine Expert
 *                         仅依赖 IEC 61131-3 算术运算符与 ABS，零厂商私有库
 * 功能描述 (Function)   : 带上下限的原地递减饱和（FC 形态）：把 VAR_IN_OUT 引脚 fX 原地
 *                         −1.0（步进常量 DL_SDEC_STEP），结果低于下限 fMin 则饱和到 fMin，
 *                         高于上限 fMax 则压回 fMax。与 FC_DL_SaturateIncr 严格对称，
 *                         共用 E_DL_SaturateErr 枚举（属主为递增件）。
 *                         **原地语义**：写回点唯一（各分支末端），返回 FALSE 的所有出口
 *                         均不写 fX，保证「失败不推进」。
 * 接口     (Interface)  : VAR_IN_OUT fX 被递减的量（本件原地更新）[工程单位]；
 *                         输入 fMin 下限、fMax 上限（有效域 fMin ≤ fMax）[工程单位]；
 *                         输出 fY 递减后值（镜像 fX）[工程单位]、bSaturated 本拍是否饱和、
 *                         eErrCode（E_DL_SaturateErr，引用不重声明）；返回值 = 递减已生效标志。
 * 边界     (Boundary)   : ① fMin > fMax → 故障级 eBadLimit，fX 不写回。
 *                         ② 任一入参非有限 → 故障级 eNonFinite，fX 不写回。
 *                         ③ fX − 1 溢出为非有限 → 故障级 eNonFinite，fX 不写回。
 *                         ④ 下限饱和与上限压回为两个独立分支、两个独立码值（R190 归因唯一）。
 *                         ⑤ 容差 DL_SDEC_EPS（1E-6）用于限值判定，禁浮点判等。
 *                         ⑥ 零全局耦合（无 GVL / VAR_EXTERNAL / 物理地址）。
 * 码表     (Codes)      : 本件不占用全局数字码位（R297 零码位范式）；出口复用
 *                         E_DL_SaturateErr，属主 FC_DL_SaturateIncr.st，本件只引用。
 * 分工声明 (Scope)      : 递增同族件为 FC_DL_SaturateIncr（枚举属主）；整数类限位递减
 *                         归 FC_DL_ClampDintChk 与 FC_DL_BcdDecrementByte。
 * 归属     (Ownership)  : E_DL_SaturateErr 归属 FC_DL_SaturateIncr.st，本件只引用不重声明。
 * 红线自检 (Redline)    : R1 ✓ 零 GVL ｜ R2 ✓ 零 %I/%Q ｜ R3 ✓ 纯 IEC ｜ R4 ✓ 非有限双判 +
 *                         上下限域闸 + 容差比较 ｜ R5 ✓ 逐行同行双语注释 ｜ R6 N/A（纯函数）
 *                         R7 N/A（无实例调用）
 * 修订历史 (Revision)   : 2026-11-23  v1.0.0  R78-B2 首版
 * 验收向量 (Acceptance) :
 *   A1 fX=4.0, fMin=0.0, fMax=10.0 → fX=3.0, fY=3.0, bSaturated=FALSE, eIncremented；
 *   A2 fX=0.0, fMin=0.0, fMax=10.0 → fX=0.0, bSaturated=TRUE, eSatLow；
 *   A3 fX=0.5, fMin=0.0, fMax=10.0 → fX=0.0, bSaturated=TRUE, eSatLow；
 *   A4 fX=10.5, fMin=0.0, fMax=10.0 → fX=10.0, bSaturated=TRUE, eSatHigh（压回上限）；
 *   A5 fX=5.0, fMin=10.0, fMax=0.0 → fX 保持 5.0, eBadLimit, 返回 FALSE。
 *============================================================================*)

FUNCTION FC_DL_SaturateDecr : BOOL
VAR_IN_OUT
    fX : LREAL;      // 被原地递减的量，成功时本件写回新值 [工程单位] / Value decremented in place, written back on success
END_VAR
VAR_INPUT
    fMin : LREAL;    // 下限 [工程单位] / Low limit in engineering unit
    fMax : LREAL;    // 上限，有效域 ≥ fMin [工程单位] / High limit in engineering unit, valid domain >= fMin
END_VAR
VAR_OUTPUT
    fY         : LREAL;             // 递减后值（镜像 fX）[工程单位] / Decremented value, mirror of fX
    bSaturated : BOOL;              // 本拍是否发生饱和 [-] / Saturation flag of this scan
    eErrCode   : E_DL_SaturateErr;  // 出口码（引用递增件属主枚举）[-] / Outlet code referencing the owner enum
END_VAR
VAR
    _bBadX   : BOOL;   // fX 非有限标志 [-] / Non-finite flag of fX
    _bBadMin : BOOL;   // fMin 非有限标志 [-] / Non-finite flag of fMin
    _bBadMax : BOOL;   // fMax 非有限标志 [-] / Non-finite flag of fMax
    _fNext   : LREAL;  // 裸递减结果 = fX − 步进 [工程单位] / Raw decremented value before saturation
END_VAR
VAR CONSTANT
    DL_SDEC_ZERO : LREAL := 0.0;     // 零基准 [-] / Zero base
    DL_SDEC_ONE  : LREAL := 1.0;     // 递减步进常量 [-] / Decrement step constant
    DL_SDEC_EPS  : LREAL := 1.0E-6;  // 限值比较容差 [-] / Limit comparison tolerance
END_VAR

(* —— 段 0：出口预置安全侧 —— *)
FC_DL_SaturateDecr := FALSE;                         // 返回值预置未生效 / Return preset not applied
fY         := fX;                                    // 镜像出口取原值（失败不推进）/ Mirror keeps the original value on failure
bSaturated := FALSE;                                 // 饱和标志预清（单拍位统一预置）/ Single-shot flag preset
eErrCode   := E_DL_SaturateErr.eNonFinite;           // 预置最严码 / Preset strictest code

(* —— 段 1：入参非有限闸（R272 全量枚举 fX / fMin / fMax） —— *)
_bBadX   := (fX <> fX) OR ((fX - fX) <> DL_SDEC_ZERO);                       // 被递减量非有限 / Value non-finite
_bBadMin := (fMin <> fMin) OR ((fMin - fMin) <> DL_SDEC_ZERO);               // 下限非有限 / Low limit non-finite
_bBadMax := (fMax <> fMax) OR ((fMax - fMax) <> DL_SDEC_ZERO);               // 上限非有限 / High limit non-finite
IF _bBadX OR _bBadMin OR _bBadMax THEN
    RETURN;                                          // 故障出口：fX 不写回 / Fault exit, fX not written
END_IF

(* —— 段 2：上下限域闸（倒置即组态缺陷，拒绝且不写回） —— *)
IF fMin > (fMax + DL_SDEC_EPS) THEN
    eErrCode := E_DL_SaturateErr.eBadLimit;          // 故障级码 / Fault-level code
    RETURN;                                          // 返回 FALSE / Fault exit
END_IF

(* —— 段 3：裸递减与溢出复检 —— *)
_fNext := fX - DL_SDEC_ONE;                          // 裸递减 / Raw decrement
IF (_fNext <> _fNext) OR ((_fNext - _fNext) <> DL_SDEC_ZERO) THEN
    eErrCode := E_DL_SaturateErr.eNonFinite;         // 故障级码：溢出为非有限 / Fault: overflow to non-finite
    RETURN;                                          // 返回 FALSE，fX 不写回 / Fault exit
END_IF

(* —— 段 4：下限饱和（独立分支 + 独立码值，R190） —— *)
IF _fNext < fMin THEN
    fY         := fMin;                              // 饱和到下限 / Saturate at the low limit
    fX         := fMin;                              // 原地写回（唯一写回点）/ Single write-back point
    bSaturated := TRUE;                              // 饱和标志 / Saturation flag
    eErrCode   := E_DL_SaturateErr.eSatLow;          // 信息级：下限饱和 / Info: saturated low
    FC_DL_SaturateDecr := TRUE;                      // 递减已生效（饱和后值）/ Decrement applied with saturation
    RETURN;
END_IF

(* —— 段 5：上限压回（独立分支 + 独立码值，R190） —— *)
IF _fNext > fMax THEN
    fY         := fMax;                              // 压回到上限 / Clamp back to the high limit
    fX         := fMax;                              // 原地写回（唯一写回点）/ Single write-back point
    bSaturated := TRUE;                              // 饱和标志 / Saturation flag
    eErrCode   := E_DL_SaturateErr.eSatHigh;         // 信息级：上限饱和 / Info: saturated high
    FC_DL_SaturateDecr := TRUE;                      // 递减已生效（压回后值）/ Decrement applied with clamp
    RETURN;
END_IF

(* —— 段 6：限内正常推进 —— *)
fY         := _fNext;                                // 正常推进结果 / Normal decremented value
fX         := _fNext;                                // 原地写回（唯一写回点）/ Single write-back point
bSaturated := FALSE;                                 // 未饱和 / Not saturated
eErrCode   := E_DL_SaturateErr.eIncremented;         // 信息级：限内推进（共用成员）/ Info: advanced within limits
FC_DL_SaturateDecr := TRUE;                          // 递减已生效 / Decrement applied
END_FUNCTION

(* ---- FC_DL_SearchMinMax.st ---- *)
(*==============================================================================
 * 组件名称 (Component)  : FC_DL_SearchMinMax
 * 所属子库 (Sublibrary) : DL_MathData
 * 当前版本 (Version)    : 1.0.0
 * 组件分类 (Category)   : 函数（FUNCTION）· 纯函数 · 数组极值与索引同出
 * 兼容性   (Platform)   : CODESYS 3.5 / TwinCAT 3 / 汇川 InoProShop / Schneider
 *                         Machine Expert；仅用 ABS / MIN / MAX 等标准算子
 * 功能描述 (Function)   : 在注入数组的前 nCount 个元素中一次单遍扫描，同时求
 *                         最小值、最大值及其索引（可选首个命中或末次命中），
 *                         并统计被跳过的非有限值（NaN 与超大值）个数。用于
 *                         批次数据极值分析、多路温度最高点定位、传感器阵列
 *                         故障点筛查、配方曲线包络提取。
 * 与既有件边界 (Boundary): FB_DL_SignalStatistics 是流式窗口统计（有状态、
 *                         含均值方差）；FB_DL_PeakDetector 是时域峰值跟踪
 *                         （带衰减与事件）；本件是静态数组一次性扫描（纯函数、
 *                         无状态），只出极值与索引，不做任何时间维度处理。
 * 设计要点 (Key notes)  : ① 单遍扫描：一趟循环同时出极值与索引，不做两次
 *                           遍历（大数组下 O(2N) 与 O(N) 的差别会被任务周期
 *                           放大）；
 *                         ② 首命中用严格比较、末命中用非严格比较，不以
 *                           MODE 参数区分（单一布尔策略开关，语义单一，
 *                           不构成多职责巨无霸块）；
 *                         ③ 非有限值过滤不依赖厂商 ISNAN 函数：用「NaN 不等于
 *                           自身」这一 IEEE 754 可移植判据，配合绝对值超
 *                           1E300 兜底无穷大，两条件任一成立即跳过；
 *                         ④ 全量非有限时返回 FALSE 并置故障级码，绝不用 0 冒充
 *                           有效极值（否则上层会把「无数据」当成「最小值 0」）；
 *                         ⑤ 数组上界必须用钳位后的局部变量，禁止直接用入参
 *                           nCount 当 FOR 上界（越界访问是 PLC 上最典型的
 *                           内存踩踏来源）。
 * 开源溯源 (Origin)     : lgf-math。参考 LGF（Libre Graphical Framework）公开
 *                         函数库「Math」分类下 SearchMinMax 系列的四个类型
 *                         变体（LReal / DInt / UDInt / 通用）所体现的功能
 *                         分类与参数域（数据体 + 个数 + 极值 + 索引 的参数
 *                         形态），只借分类、参数域与命名习惯；本件只做 LREAL
 *                         主线，其余类型变体按库内「数据类型重载」规则另立块，
 *                         不塞进 MODE 参数。算法与实现 100% 自有 clean-room，
 *                         不构成衍生作品。
 * 依赖     (Depends)    : 无 DL_ 内部依赖；无标准库功能块依赖
 * 故障码表 (Error codes):
 *   16#0001_0119【信息级】计数越界（小于 1 早退；大于上限则钳位后继续）
 *   16#0001_011A【信息级】检测到非有限值并已跳过，个数见 nSkipCnt
 *   16#0001_0217【故障级】全量非有限，无有效极值，返回 FALSE
 * 验收向量 (Acceptance) :
 *   V1 数据 3.5 / -2.0 / 9.0 / -2.0，个数 4，首命中 → 最小 -2.0 于索引 1，
 *      最大 9.0 于索引 2
 *   V2 同上改末次命中 → 最小 -2.0 于索引 3
 *   V3 数据 1.0 / NaN / 1.0 → 跳过 1 个、有效 2 个、全等标志 TRUE、码含 011A
 *   V4 个数 0 → 返回 FALSE、码 0119、两个索引均为 -1
 *   V5 个数 300（超 256）→ 只扫前 256 个、码 0119、返回 TRUE
 * 红线自检 (Redline)    : R1 零全局变量表与外部变量引用 ｜ R2 零物理地址直写
 *                         R3 纯 IEC 61131-3 ｜ R4 索引先钳位后访问、浮点比较
 *                         用容差、NaN 判据有注释豁免说明 ｜ R5 全变量中英双语
 *                         同行注释 ｜ R6 N/A（纯函数无状态机）｜ R7 N/A（无实例）
 * 修订历史 (Revision)   :
 *   2026-11-15  v1.0.0  首版入库（Round 10 · Level 1 数学族回补）
 *============================================================================*)

FUNCTION FC_DL_SearchMinMax : BOOL
VAR_INPUT
    nCount   : DINT := 0;        // 参与扫描的元素个数，有效域 1 到 DL_SMM_MAX [个] / Number of elements to scan, valid 1 to DL_SMM_MAX
    bLastHit : BOOL := FALSE;    // TRUE = 索引取末次命中，FALSE = 取首个命中（默认）[-] / TRUE selects the last hit, FALSE the first hit
END_VAR
VAR_IN_OUT
    afData   : ARRAY[0..255] OF LREAL;  // 扫描数据体，调用方持有并注入，上界 255 与 DL_SMM_MAX 保持一致 [工程单位] / Scanned data array, bound 255 kept in sync with DL_SMM_MAX
END_VAR
VAR_OUTPUT
    fMin      : LREAL;       // 最小值，无有效数据时为 0.0 [工程单位随应用] / Minimum value, 0.0 when no valid element
    fMax      : LREAL;       // 最大值，无有效数据时为 0.0 [工程单位随应用] / Maximum value, 0.0 when no valid element
    nMinIdx   : DINT := -1;  // 最小值索引，未找到为 -1 [元素下标] / Index of the minimum, -1 when not found
    nMaxIdx   : DINT := -1;  // 最大值索引，未找到为 -1 [元素下标] / Index of the maximum, -1 when not found
    nValidCnt : DINT;        // 实际参与比较的有效元素数 [个] / Number of elements actually compared
    nSkipCnt  : DINT;        // 因非有限值被跳过的元素数 [个] / Number of skipped non-finite elements
    bFlat     : BOOL;        // 全等标志，fMin 与 fMax 在容差内相等 [-] / TRUE when the minimum equals the maximum within tolerance
    uErrorId  : UDINT;       // 事件码，0 = 无事件 / Event code, 0 = no event
END_VAR
VAR
    i            : DINT;     // 循环索引，域 0 到钳位后个数减 1 [元素下标] / Loop index, 0 to clamped count minus one
    nCountClamp  : DINT;     // 钳位后的扫描个数，FOR 上界只许用本变量 [个] / Clamped scan count, the only legal FOR upper bound
    fValue       : LREAL;    // 当前元素值副本，避免在比较中重复取数组 [工程单位] / Current element value copy
    bFinite      : BOOL;     // 当前元素是否有限（非 NaN 且非超大幅值）[-] / TRUE when the current element is finite
END_VAR
VAR CONSTANT
    DL_SMM_MAX   : DINT  := 256;      // 数组上限，与形参上界 255 保持一致 [元素] / Array upper bound, kept in sync with the formal bound
    DL_SMM_MIN   : DINT  := 1;        // 最小扫描个数，0 与负数一律视为非法 [个] / Minimum legal scan count
    DL_FLOAT_EPS : LREAL := 1.0E-9;   // 浮点比较容差，用于全等判定 [-] / Float comparison tolerance for the flat test
    DL_BIG       : LREAL := 1.0E300;  // 超大值兜底门限，用于识别无穷大与溢出 [-] / Magnitude guard used to catch infinities
END_VAR

(*------------------------------------------------------------------------------
 * 段 1｜输出与返回值预置：早退路径必须给出确定的 0 与 -1
 *      Pre-set outputs: deterministic zeros and minus one on every early exit
 *-----------------------------------------------------------------------------*)
FC_DL_SearchMinMax := FALSE;
fMin      := 0.0;
fMax      := 0.0;
nMinIdx   := -1;
nMaxIdx   := -1;
nValidCnt := 0;
nSkipCnt  := 0;
bFlat     := FALSE;
uErrorId  := 16#0000_0000;

(*------------------------------------------------------------------------------
 * 段 2｜计数域校验（边界 B1）：小于 1 直接早退，大于上限钳位后继续
 *      Count domain check: below one exits early, above the bound is clamped
 *      钳位而不报错退出的理由：现场宁可算出前 256 个的极值，也不要拿不到数
 *-----------------------------------------------------------------------------*)
IF nCount < DL_SMM_MIN THEN
    uErrorId := 16#0001_0119;   // 计数非法（小于 1），无有效极值
    RETURN;
END_IF

nCountClamp := nCount;
IF nCount > DL_SMM_MAX THEN
    nCountClamp := DL_SMM_MAX;  // 只扫前 DL_SMM_MAX 个，绝不越界
    uErrorId    := 16#0001_0119;
END_IF

(*------------------------------------------------------------------------------
 * 段 3｜单遍扫描：过滤非有限值，同时维护极值与索引
 *      Single pass: filter non-finite values while tracking extremes and indices
 *      NaN 判据：fValue 不等于 fValue 在 IEEE 754 下恒为 TRUE（NaN 不等于自身），
 *      这是唯一可移植的 NaN 检测手段，不依赖任何厂商 ISNAN 函数；
 *      绝对值超过 1E300 视为无穷大或数值溢出，一并跳过。
 *-----------------------------------------------------------------------------*)
FOR i := 0 TO (nCountClamp - 1) DO
    fValue := afData[i];

    IF (fValue <> fValue) OR (ABS(fValue) > DL_BIG) THEN
        bFinite := FALSE;
    ELSE
        bFinite := TRUE;
    END_IF

    IF NOT bFinite THEN
        nSkipCnt := nSkipCnt + 1;               // 非有限值：跳过，不参与比较
    ELSE
        IF nValidCnt = 0 THEN
            fMin     := fValue;                 // 首个有效元素直接作为初值
            fMax     := fValue;
            nMinIdx  := i;
            nMaxIdx  := i;
        ELSE
            IF bLastHit THEN
                IF fValue <= fMin THEN          // 末命中：等值也替换索引
                    fMin    := fValue;
                    nMinIdx := i;
                END_IF
                IF fValue >= fMax THEN
                    fMax    := fValue;
                    nMaxIdx := i;
                END_IF
            ELSE
                IF fValue < fMin THEN           // 首命中：等值不替换索引
                    fMin    := fValue;
                    nMinIdx := i;
                END_IF
                IF fValue > fMax THEN
                    fMax    := fValue;
                    nMaxIdx := i;
                END_IF
            END_IF
        END_IF
        nValidCnt := nValidCnt + 1;
    END_IF
END_FOR

(*------------------------------------------------------------------------------
 * 段 4｜全量非有限兜底（边界 B2）：无有效元素时绝不返回 0 冒充极值
 *      All non-finite fallback: never report zero as a valid extreme
 *-----------------------------------------------------------------------------*)
IF nValidCnt < 1 THEN
    fMin     := 0.0;
    fMax     := 0.0;
    nMinIdx  := -1;
    nMaxIdx  := -1;
    uErrorId := 16#0001_0217;   // 故障级：无有效极值
    FC_DL_SearchMinMax := FALSE;
    RETURN;
END_IF

(*------------------------------------------------------------------------------
 * 段 5｜全等判定（浮点禁用判等）：用容差比较代替相等比较
 *      Flat detection with a tolerance compare instead of an equality compare
 *-----------------------------------------------------------------------------*)
IF ABS(fMax - fMin) < DL_FLOAT_EPS THEN
    bFlat := TRUE;
ELSE
    bFlat := FALSE;
END_IF

(*------------------------------------------------------------------------------
 * 段 6｜事件码收口：数据质量问题优先于计数钳位事件
 *      Error code close-out: data quality outranks the count clamp event
 *-----------------------------------------------------------------------------*)
IF nSkipCnt > 0 THEN
    uErrorId := 16#0001_011A;   // 信息级：存在被跳过的非有限值
END_IF

FC_DL_SearchMinMax := TRUE;
END_FUNCTION

(* ---- FC_DL_SearchMinMaxDint.st ---- *)
(*
  ==================================================================
  组件名 Component  : FC_DL_SearchMinMaxDint
  分类   Category   : DL_MathData
  复杂度 Complexity  : 低
  版本   Version    : 1.0.0
  功能   Purpose    : DINT 域数组单遍扫描求最小值/最大值与双索引同出。前 nCount
                      个元素有效，一次循环同时出 nMin/nMax 与 uMinIdx/uMaxIdx
                      （首命中口径），无效哨兵按开关跳过并计数。
  来源   Source     : t2-1-lgf-math（LGF Math 极值检索族 DINT 变体）
  溯源   Origin     : 极值检索属公开数学语义，clean-room 自研实现，未复制 LGF
                      或任何厂商私有库源码。
  平台   Platform   : 纯 IEC 61131-3（仅 FOR / 比较 / DINT_TO_UDINT），
                      CODESYS / TwinCAT / InoProShop / Machine Expert 通用
  分工声明 Split     : 与 FC_DL_SearchMinMax（LREAL 属主）互引——后者管 LREAL
                      域并以 x <> x 剔除 NaN；本件为 DINT 域重载，只做整数极值，
                      不做浮点有限性判据。与 FC_DL_SearchMinMaxUdint 同批成对，
                      共用同一规格向量表、码位段同带连号。
  作者   Author     : 道莅代码库 · PLC 编程专家（R60）
  ------------------------------------------------------------------
  边界 Boundary     :
                      一 扫描个数钳位 1..4096，钳位置信息级码；
                      二 无效样本域：DINT 域无 NaN（LREAL 属主用 x <> x 判据），
                         本件无效量定义为哨兵 DL_SMM_INVALID（等于 DINT 最小值
                         位型 16#8000_0000），仅当 bIgnoreInvalid 为真时跳过；
                      三 全量无效时不返回 0 号位「伪极值」——bValid = FALSE 且
                         两个索引回 0，由调用方按 bValid 判别（沿 LREAL 属主纪律）；
                      四 索引写出前已证在 [0, nUse-1] 内，回钳后不再复判越界（R241）；
                      五 无状态纯函数：每次调用局部量一律段 1 显式预置（R254）。
  接口偏离声明       : 派单示意 fMin/fMax（浮点命名），DINT 输出按 R265 命名-类型
                      一致性落为 nMin/nMax，语义与引脚数一字不减。
  错误码   Codes    :
    16#0001_0601【信息级】计数越界已钳位（<1 早退，>4096 钳位续扫）
    16#0001_0602【信息级】无效哨兵样本已跳过，个数见 nSkipCnt
    16#0001_0603【故障级】全量无效，无有效极值，bValid = FALSE
  验收   Acceptance :
    算法已证（脚本）：未跑 ｜ 编译器已证（三平台）：未跑
    V1 数据 5 / -3 / 9 / -3，个数 4 → nMin=-3 于索引 1，nMax=9 于索引 2
    V2 数据 7 / 7 / 7 → nMin=nMax=7，双索引均 0（首命中）
    V3 哨兵 16#8000_0000 夹在有效值间，bIgnoreInvalid 真 → 跳过 1 个，码含 0602
    V4 个数 0 → bValid=FALSE、码 0601、双索引 0
    V5 全为哨兵且 bIgnoreInvalid 真 → bValid=FALSE、码 0603
  修订记录 Revision  :
    2026-11-21  v1.0.0  R60 首版（批 1 · 序号 1）
  ==================================================================
*)
FUNCTION FC_DL_SearchMinMaxDint : BOOL
VAR_IN_OUT
    aValues : ARRAY[0..4095] OF DINT; // 待扫描数组 [工程计数]，前 nCount 个有效 / the scanned array, the first nCount entries valid
END_VAR
VAR_INPUT
    nCount         : DINT; // 有效样本数 [个]，钳位 1..4096 / the valid sample count, clamped to one through four thousand ninety six
    bIgnoreInvalid : BOOL; // 是否跳过无效哨兵值 [-] / whether the invalid sentinel entries are skipped
END_VAR
VAR_OUTPUT
    nMin     : DINT;  // 最小值 [工程计数]，无有效样本时为 0 / the minimum value, zero when no valid sample
    nMax     : DINT;  // 最大值 [工程计数]，无有效样本时为 0 / the maximum value, zero when no valid sample
    uMinIdx  : UDINT; // 最小值所在下标 [下标]，无有效样本时为 0 / the minimum index, zero when no valid sample
    uMaxIdx  : UDINT; // 最大值所在下标 [下标]，无有效样本时为 0 / the maximum index, zero when no valid sample
    nSkipCnt : UDINT; // 被跳过的无效哨兵个数 [个] / the skipped invalid sentinel count
    bValid   : BOOL;  // 结果是否有效（全量无效时为假）[-] / the result validity flag
    eErr     : UDINT; // 错误码，0 = 正常 / the error code, zero is ok
    bError   : BOOL;  // 错误标志，eErr 非 0 时为真 / the error flag, true when eErr is nonzero
END_VAR
VAR
    nI      : DINT;  // 扫描索引 [下标] / the scan index
    nUse    : DINT;  // 钳位后的扫描个数 [个] / the clamped scan count
    nSeen   : DINT;  // 已见有效样本数 [个] / the seen valid sample count
    nV      : DINT;  // 当前样本工作副本 [工程计数] / the current sample working copy
    bHave   : BOOL;  // 已取得首个有效样本 [-] / the first valid sample taken flag
    bClamp  : BOOL;  // 钳位发生标记 [-] / the clamp happened flag
END_VAR
VAR CONSTANT
    DL_SMM_DMAX      : DINT := 4096;               // 扫描个数上界 [个]，与数组容量一致 / the scan count bound aligned with the array capacity
    DL_SMM_INVALID   : DINT := -16#7FFF_FFFF - 1;  // 无效哨兵，等于 DINT 最小位型 16#8000_0000（禁用超域字面量写法）/ the invalid sentinel equal to the DINT minimum bit pattern
END_VAR

// 段 1｜返回值与错误状态预置安全值（四段式第一段，R45）+ 局部量显式预置（R254）/ segment 1, the preset of the return, the codes and the local guards
FC_DL_SearchMinMaxDint := FALSE; // 返回值预置假 / preset the return false
nMin := 0; // 最小值预置零 / preset the minimum zero
nMax := 0; // 最大值预置零 / preset the maximum zero
uMinIdx := 0; // 最小索引预置零 / preset the minimum index zero
uMaxIdx := 0; // 最大索引预置零 / preset the maximum index zero
nSkipCnt := 0; // 跳过计数预置零 / preset the skipped count zero
bValid := FALSE; // 有效标志预置假（无有效样本前不宣称有效）/ preset the validity false
eErr := 16#0000_0000; // 错误码预置正常 / preset the code to ok
bError := FALSE; // 错误标志预置假 / preset the error flag false
nUse := 0; // 扫描个数预置零 / preset the scan count zero
nSeen := 0; // 有效样本数预置零 / preset the seen count zero
nV := 0; // 样本工作副本预置零 / preset the sample copy zero
bHave := FALSE; // 首样本标志预置假 / preset the first sample flag false
bClamp := FALSE; // 钳位标记预置假 / preset the clamp flag false

// 段 2｜扫描个数域闸（下界早退 + 上界钳位，边界一）/ segment 2, the scan count domain gate
IF nCount < 1 THEN // 低于下界，无样本可扫 / below the floor, nothing to scan
    eErr := 16#0001_0601; // 信息级：计数越界已钳位 / informational, the count clamped
    bError := TRUE; // 置错误标志（信息级随事件置位惯例）/ raise the error flag
    RETURN; // 早退：bValid 保持 FALSE，双索引保持 0 / early return with the validity false
END_IF
nUse := nCount; // 域内接管 / take the count inside the domain
IF nUse > DL_SMM_DMAX THEN // 高于上界 / above the bound
    nUse := DL_SMM_DMAX; // 钳到数组容量 / clamp to the array capacity
    bClamp := TRUE; // 置钳位标记 / raise the clamp flag
END_IF
IF bClamp THEN // 钳位发生时置信息级 / raise the informational code on a clamp
    eErr := 16#0001_0601; // 信息级：计数越界已钳位 / informational, the count clamped
    bError := TRUE; // 置错误标志 / raise the error flag
END_IF

// 段 3｜单遍扫描：首命中取极小与极大，索引与值同源写出（边界四）/ segment 3, the single pass scan with the first hit rule
FOR nI := 0 TO nUse - 1 DO // 有界循环（nUse 已钳 ≤4096）/ the bounded loop
    nV := aValues[nI]; // 取样本（索引已证在数组界内）/ take the sample, the index proven inside the bounds
    IF bIgnoreInvalid AND (nV = DL_SMM_INVALID) THEN // 无效哨兵且开关为真 / an invalid sentinel with the switch true
        nSkipCnt := nSkipCnt + 1; // 跳过计数推进 / advance the skipped count
    ELSE // 有效样本参与极值 / a valid sample participates
        nSeen := nSeen + 1; // 有效样本数推进 / advance the seen count
        IF NOT bHave THEN // 首个有效样本：双向装填 / the first valid sample seeds both sides
            nMin := nV; // 最小值装填 / seed the minimum
            nMax := nV; // 最大值装填 / seed the maximum
            uMinIdx := DINT_TO_UDINT(nI); // 最小索引装填 / seed the minimum index
            uMaxIdx := DINT_TO_UDINT(nI); // 最大索引装填 / seed the maximum index
            bHave := TRUE; // 置首样本标志 / raise the first sample flag
        ELSE // 后续样本比较（首命中用严格比较，不覆盖等值）/ the later samples, strict compare keeps the first hit
            IF nV < nMin THEN // 新极小 / a new minimum
                nMin := nV; // 更新最小值 / update the minimum
                uMinIdx := DINT_TO_UDINT(nI); // 更新最小索引（与值同源）/ update the minimum index from the same source
            ELSIF nV > nMax THEN // 新极大（nV ≥ nMin 前提下判极大即可，单调序自证）/ a new maximum, proven since nV is not below the minimum
                nMax := nV; // 更新最大值 / update the maximum
                uMaxIdx := DINT_TO_UDINT(nI); // 更新最大索引（与值同源）/ update the maximum index from the same source
            END_IF
        END_IF
    END_IF
END_FOR

// 段 4｜结果复检兜底：全量无效判故障，信息级与故障级不共码（R258 三件套）/ segment 4, the result recheck
IF (nSeen > 0) AND (nSkipCnt > 0) AND (eErr = 16#0000_0000) THEN // 部分跳过且无先发事件 / a partial skip with no earlier event
    eErr := 16#0001_0602; // 信息级：无效哨兵样本已跳过 / informational, the invalid sentinels skipped
    bError := TRUE; // 置错误标志 / raise the error flag
END_IF
IF nSeen < 1 THEN // 无有效样本 / no valid sample
    eErr := 16#0001_0603; // 故障级：全量无效，无有效极值 / fault grade, no valid extremum
    bError := TRUE; // 置错误标志（R45 配对）/ raise the error flag, paired with the fault code
    bValid := FALSE; // 结果不可用 / the result void
    nMin := 0; // 双极值回安全值 / both extrema back to the safe zero
    nMax := 0; // 双极值回安全值 / both extrema back to the safe zero
    uMinIdx := 0; // 索引回 0（不冒充 0 号位极值，边界三）/ the index back to zero, not posing as the entry zero
    uMaxIdx := 0; // 索引回 0（不冒充 0 号位极值，边界三）/ the index back to zero, not posing as the entry zero
ELSE // 有有效样本 / with valid samples
    bValid := TRUE; // 结果有效 / the result is valid
    FC_DL_SearchMinMaxDint := TRUE; // 返回成功 / return success
END_IF
END_FUNCTION
